(* IEC 61131-3 sources: daoli-st-library/DL_Base (part 20) *)

(* ---- FB_DL_PresetCounterSat.st ---- *)
(*==============================================================================
 * 组件名称 (Component)  : FB_DL_PresetCounterSat
 * 所属子库 (Sublibrary) : DL_Base
 * 当前版本 (Version)    : 1.0.1
 * 分类     (Category)   : 计数功能块（Function Block · Counter）
 * 兼容性   (Platform)   : CODESYS 3.5 / TwinCAT 3 / 汇川 InoProShop / Machine Expert
 *                         仅依赖 Standard.library（R_TRIG），零厂商方言
 * 功能简介 (Function)   : 带饱和预设计数器：上/下双向计数（上升沿生效），
 *                         到达上限（nPreset）或下限（nLowLimit）饱和不回绕
 *                         ——上计数在 nCount >= nPreset 时拒绝递增并保持
 *                         bSatHigh，下计数在 nCount <= nLowLimit 时拒绝递减
 *                         并保持 bSatLow。到达上限输出保持型完成标志 bDone
 *                         与单拍阈值事件 bThreshold（首次到达一拍脉冲，遵循
 *                         R25 单拍标志生命周期三律）。装载 bLoad 优先级最高，
 *                         复位 bReset 次之，同拍双计数互相抵消不偏置任何方向。
 *                         与已入库 FB_DL_EventCounter（回绕 + 比较输出通用
 *                         事件计数）、FB_DL_ModuloCounter（取模工位索引）
 *                         职责分离——本块是饱和计数（批次计数 / 托盘满载
 *                         场景），越界语义固定为钳位停走。
 * 开源溯源 (Origin)     : 原创实现（参考 LGF 库 Counter 计数器分类的功能域
 *                         与参数域，来源标签 lgf-counter），饱和计数语义为
 *                         公开计数器行为域，仅借分类/参数域/命名，clean-room
 *                         实现，未复制任何厂商私有库源码，不构成衍生作品。
 * 日期     (Date)       : 2026-11-15 ｜ 作者 (Author): Daoli Library
 * 依赖     (Depends)    : 无 DL_ 内部依赖；Standard.library: R_TRIG
 *
 *------------------------------------------------------------------------------
 * 【引脚契约 / Pin contract】
 *   输入 bCountUp   : BOOL — 上计数脉冲输入，上升沿 +1；
 *   输入 bCountDown : BOOL — 下计数脉冲输入，上升沿 -1；
 *   输入 bLoad      : BOOL — 装载预设值，上升沿生效（优先级最高）；
 *   输入 nPreset    : DINT — 上限预设值 [个]，>= nLowLimit，默认 100；
 *   输入 nLowLimit  : DINT — 下限预设值 [个]，<= nPreset，默认 0；
 *   输入 bReset     : BOOL — 复位到下限，上升沿生效（次优先级，兼故障解除）；
 *   输出 nCount     : DINT — 当前计数值 [个]，饱和域 [nLowLimit, nPreset]；
 *   输出 bSatHigh   : BOOL — 已达上限饱和（保持型，逐拍重算）；
 *   输出 bSatLow    : BOOL — 已达下限饱和（保持型，逐拍重算）；
 *   输出 bDone      : BOOL — 计数到达上限（保持型，逐拍重算）；
 *   输出 bThreshold : BOOL — 首次到达上限单拍脉冲（R25 三律）；
 *   输出 uErrorId   : UDINT — 故障码，0 = 无故障。
 *
 * 【优先级序 / Priority order（写死防歧义）】
 *   参数故障锁存 > 装载（bLoad 沿）> 复位（bReset 沿）> 同拍双计数抵消
 *   （计数值不变，不偏置任何方向）> 单向上计数 > 单向下计数 > 保持。
 *   同拍装载与计数脉冲：装载覆盖计数（计数脉冲被吞，不补发不记账）。
 *   同拍装载与复位：装载优先（覆盖复位到下限的行为）。
 *
 * 【饱和语义 / Saturation semantics（写死防误解）】
 *   上饱和：nCount = nPreset 时再收上计数沿 → 计数值保持 nPreset 不回绕、
 *           不取模，bSatHigh 保持 TRUE，脉冲被吞不置任何事件码（饱和本身
 *           是正常工况语义而非故障，上层以 bSatHigh/bDone 感知）；
 *   下饱和：nCount = nLowLimit 时再收下计数沿 → 保持 nLowLimit，bSatLow
 *           保持 TRUE，脉冲同样被吞；
 *   与 FB_DL_EventCounter 的 bWrap = FALSE 饱和模式语义一致但本块无回绕
 *   选项——批次/满载场景回绕是危险行为，设计上直接删除该自由度。
 *
 * 【bThreshold 单拍 R25 三律落地 / One-shot pulse lifecycle】
 *   置位律：仅「本拍到达上限 AND 上拍未在限」的扫描拍置 TRUE
 *           （bReached 为边沿基准，单一来源，仅由计数出口单点推导）；
 *   自清律：bThreshold 每拍预清 FALSE，无到达沿自动回落，不锁存；
 *   基准律：bReached 每拍在计数出口后单点刷新为 (nCount >= nPreset)，
 *           无第二份镜像状态；故障拍强制 bReached := FALSE，故障解除后
 *           再次到达会重新给出一拍脉冲（诊断链可见）。
 *
 * 【边界防错清单 / Boundary guard list】
 *   B1 nPreset < nLowLimit → 参数非法故障锁存 16#0001_0212：计数值强制钳到
 *      nLowLimit，计数/装载全部冻结，仅 bReset 上升沿解除（R15：故障级
 *      锁存仅解除路径清码）；解除后首次满足条件重新计数；
 *   B2 先判界后加减：上计数前判 nCount >= nPreset、下计数前判
 *      nCount <= nLowLimit，杜绝 DINT 极值 +1/-1 回绕穿透判据；
 *   B3 同拍 bCountUp/bCountDown 同时有效 → 计数不变（不偏置任何方向）；
 *   B4 装载值即 nPreset 引脚现值（装载拍实时采样，非缓存旧值）；
 *   B5 bReset 上升沿把计数值直接置 nLowLimit 并同时清除故障锁存。
 *
 * 【调用示例 / Call example】
 *   「托盘满载计数：装满 100 件给满托信号，人工换托后复位」
 *   fbPalletCnt(bCountUp := bPartInFeed, bCountDown := bPartRejectOut,
 *               bLoad := FALSE, nPreset := 100, nLowLimit := 0,
 *               bReset := bPalletChanged, nCount => nPalletCount,
 *               bSatHigh => , bSatLow => , bDone => bPalletFull,
 *               bThreshold => bPalletFullPulse, uErrorId => uCntErr);
 *
 * 【平台移植注意 / Porting notes】
 *   全部运算为 DINT 整数比较与加减，先判界后运算的次序保证永不触发
 *   DINT 极值回绕，无浮点、无除法、无定时依赖，各平台行为一致。
 *
 * 【工程背景与应用场景 / Background and use cases】
 *   ① 托盘满载计数：产线件流逐件 +1，装满 nPreset 件给满托信号（bDone/
 *      bThreshold），人工换托后 bReset 清零重新计件；
 *   ② 批次计数器：批次目标 nPreset 件，剔除品经 bCountDown 回退，计数
 *      上下饱和防止误键导致的负数或超量程静默错值；
 *   ③ 收线长度/圈数计量：到达设定圈数停机收卷（饱和停走保证计数器停在
 *      满值可读，回绕式计数会让操作工无法读出实际完成量）；
 *   ④ 重复触发防护：bThreshold 单拍脉冲驱动一次性动作（满托打印/批次
 *      结束报文），保持型 bDone 驱动持续状态（满托指示灯）。
 *
 * 【保持型与单拍输出关系表 / Held vs one-shot output relation】
 *   输出          类型     置位条件                     复位条件
 *   bSatHigh     保持型   nCount >= nPreset            nCount 降回限内
 *   bSatLow      保持型   nCount <= nLowLimit          nCount 升回限内
 *   bDone        保持型   nCount >= nPreset            nCount 降回限内/故障
 *   bThreshold   单拍     首次到达拍（含装载到达）      下一拍自动回落
 *   bSatHigh 与 bDone 判据相同但语义分层：bSatHigh 描述"在限停走状态"，
 *   bDone 描述"任务完成状态"，分开输出便于上层对停走与完成做不同联锁。
 *
 * 【典型时序推演 / Typical timing walkthrough】
 *   设 nPreset = 3，nLowLimit = 0，上电 nCount = 0：
 *     拍 1 上沿 → 1；拍 2 上沿 → 2；拍 3 上沿 → 3，bDone TRUE，
 *       bThreshold 单拍 TRUE，bSatHigh TRUE；
 *     拍 4 上沿 → 保持 3（上饱和），bThreshold FALSE（无新到达沿）；
 *     拍 5 下沿 → 2，bSatHigh/bDone 回落，bThreshold 无脉冲（2 不是到达）；
 *     拍 6 上沿 → 3，bThreshold 单拍 TRUE（bReached 已回落，重新到达）；
 *     拍 7 bReset 沿 → 0，bSatLow TRUE，无脉冲；
 *   结论：bThreshold 严格对应"从限外进入上限"的每一次跃迁，同限保持
 *   与复位不触发，装载到达触发（口径与验收推演 C1~C7 一致）。
 *
 * 【参数退化域 / Degenerate parameter domains】
 *   nPreset = nLowLimit：计数域退化为单点，装载到该点后双向均饱和停走
 *   （验收推演 C7）；上电 nCount = 0 若低于下限（如 nLowLimit = 5），
 *   bSatLow 立即为 TRUE，首个下计数沿被吞直至装载/复位对齐下限——
 *   上层应在上电后先装载或复位一次，保证计数值落在合法饱和域内。
 *
 * 【同族职责分离 / Family separation】
 *   FB_DL_EventCounter：通用事件计数（回绕/饱和双模式 + 阈值比较输出）；
 *   FB_DL_ModuloCounter：取模工位索引（循环工位场景）；本块：固定饱和
 *   计数（批次满载），三者语义正交、零互相调用。
 *
 * 红线自检 (Redline)    : R1 零全局变量表/外部变量引用 ✓ ｜ R2 零物理 IO 地址 ✓
 *                         R3 纯 IEC 61131-3 标准运算 ✓ ｜ R4 先判界后运算/
 *                           故障锁存仅解除路径清码/参数钳位 ✓
 *                         R5 全变量中英双语同行注释 ✓ ｜ R6 N/A（无主状态机，
 *                           优先级 IF-ELSIF 链即状态裁决，规格豁免 ENUM）✓
 *                         R7 四个 R_TRIG 主体最前部无条件刷新 ✓ ｜ R8 界限/
 *                           码值全常量化，无魔法数 ✓
 * 验收推演 (Acceptance) :
 *   C1 单发递增链：nPreset=3, nLowLimit=0，连发 3 个上沿 → 1/2/3，第 3 拍
 *      bDone TRUE 且 bThreshold 单拍 TRUE；第 4 个上沿 → 保持 3，bSatHigh
 *      TRUE，bThreshold 无脉冲；
 *   C2 下饱和：nCount=0 时发下沿 → 保持 0，bSatLow TRUE，无事件码；
 *   C3 同拍双计数：nCount=1 时同拍上/下沿 → 保持 1，无偏置；
 *   C4 装载优先：nCount=0 时同拍 bLoad 沿 + 上沿 → nCount := nPreset，
 *      bThreshold 单拍 TRUE（首次到达），上沿被覆盖不记账；
 *   C5 复位：bCount=5 时 bReset 沿 → nCount := nLowLimit，bDone/bSatHigh
 *      回落，bThreshold 无脉冲（复位不算"到达"）；
 *   C6 参数非法：nPreset=2 < nLowLimit=5 → 故障锁存 0212，nCount 强制 5，
 *      计数冻结；bReset 沿 → 当拍解除锁存并把计数压到下限，但同一拍段 3
 *      复检参数仍非法即刻**重新锁存**（参数不修正则计数不恢复）；须先把
 *      nPreset 改为 >= nLowLimit，再给 bReset 沿才彻底解除并可重新计数
 *      （v1.0.1 终审勘误：原文"bReset 沿 → 解除，可重新计数"未写明参数前置，
 *      与"锁存置位每拍检测"的实现不符）；
 *   C7 下限装载边界：nPreset = nLowLimit = 7 → 上电 nCount=0，bSatLow TRUE；
 *      bLoad 沿 → nCount := 7，bThreshold 单拍 TRUE，此后双向均饱和停走。
 *
 * 【故障码表 / Error code table】
 *   16#0001_0212  参数非法：上限预设 nPreset < 下限预设 nLowLimit，故障级
 *                 锁存，计数冻结在 nLowLimit，仅 bReset 上升沿解除（0212
 *                 空闲，0210/0211 已被 EventCounter/ModuloCounter 登记）。
 *
 * 【设计要点 / Key notes】
 *   ① 计数值单点出口：段 4 优先级链只写 nWork，段 4 末 nCount := nWork
 *      单点回写，故障段强制钳位也只改出口，任何路径不出现第二份计数镜像，
 *      杜绝多出口读改写竞态（沿用库内 EventCounter 修复后的单点出口范式）；
 *   ② 先判界后运算：加/减算全部在边界预判之后执行，DINT 极值 +1/-1 回绕
 *      在数学上不可达（R25 家族通用防穿透写法）；
 *   ③ 故障锁存生命周期：置位（段 3 每拍检测）→ 冻结（段 4 闸门）→ 解除
 *      （仅段 2 复位沿），三段各一入口，无第三条改动路径（R15）；
 *   ④ 饱和吞脉冲不置码：饱和属正常工况语义，置码会造成诊断链噪音，
 *      上层以 bSatHigh/bSatLow 感知（与 EventCounter 溢出一拍脉冲口径
 *      不同，两块语义分层，注释在两侧各自写死）；
 *   ⑤ 事件型组件免首扫：计数由脉冲沿驱动，无连续量同步语义，按 R23
 *      不设 bInit 跟踪逻辑，上电即处于下限饱和观测态。
 *
 * 【实现选择 / Implementation choice】
 *   无主状态机（规格豁免 ENUM）：饱和计数的行为本质是「边沿事件 + 优先级
 *   裁决 + 单点出口」，用 IF-ELSIF 优先级链表达比 ENUM+CASE 更短且无空态；
 *   计数值单点出口（nCount := _nWork 后全段共享），bSatHigh/bSatLow/bDone
 *   全部由出口值逐拍重算派生，无第二份计数镜像，杜绝读改写竞态；
 *   本块为事件型计数组件，无连续量同步语义，按 R23 免首扫，不设 bInit。
 *
 * 修订历史 (Revision)   :
 *   2026-11-15  v1.0.0  首版落盘（Round 09 · 泳道 A · LGF Counter 组）
 *   2026-11-15  v1.0.1  终审勘误：验收推演 C6 补写"参数未修正时 bReset 沿当拍
 *                       重新锁存"的前置条件（原文易误读为复位即可恢复计数）；
 *                       代码行为未改动，故障码 0001_0212 复核无冲突
 *============================================================================*)
FUNCTION_BLOCK FB_DL_PresetCounterSat
VAR_INPUT
    bCountUp   : BOOL;                     // 上计数脉冲输入，上升沿 +1 / Count-up pulse input, rising edge increments
    bCountDown : BOOL;                     // 下计数脉冲输入，上升沿 -1 / Count-down pulse input, rising edge decrements
    bLoad      : BOOL;                     // 装载预设值，上升沿生效（优先级最高）/ Load preset, rising edge, top priority
    nPreset    : DINT := 100;              // 上限预设值 [个]，>= nLowLimit / Upper preset [pieces], at least nLowLimit
    nLowLimit  : DINT := 0;                // 下限预设值 [个]，<= nPreset / Lower preset [pieces], at most nPreset
    bReset     : BOOL;                     // 复位到下限，上升沿生效（兼故障解除）/ Reset to lower limit, rising edge, also releases the fault latch
END_VAR
VAR_OUTPUT
    nCount     : DINT := 0;                // 当前计数值 [个]，饱和域 [nLowLimit, nPreset] / Current count [pieces], saturated within [nLowLimit, nPreset]
    bSatHigh   : BOOL;                     // 已达上限饱和（保持型）/ Saturated at upper limit (held)
    bSatLow    : BOOL;                     // 已达下限饱和（保持型）/ Saturated at lower limit (held)
    bDone      : BOOL;                     // 计数到达上限（保持型）/ Count reached upper limit (held)
    bThreshold : BOOL;                     // 首次到达上限单拍脉冲（R25 三律）/ First-arrival one-shot pulse (R25 three rules)
    uErrorId   : UDINT;                    // 故障码，0 = 无故障 / Error code, 0 = none
END_VAR
VAR
    fbTrigUp   : R_TRIG;                   // 上计数边沿 / Count-up edge detector
    fbTrigDn   : R_TRIG;                   // 下计数边沿 / Count-down edge detector
    fbTrigLoad : R_TRIG;                   // 装载边沿 / Load edge detector
    fbTrigRst  : R_TRIG;                   // 复位边沿 / Reset edge detector
    bReached   : BOOL := FALSE;            // 内部到达标志（阈值事件边沿基准，单一来源）/ Internal reached flag (threshold edge baseline, single source)
    bFaultLatch: BOOL;                     // 参数非法故障锁存（仅复位沿解除）/ Invalid-parameter fault latch (released only by reset edge)
    nWork      : DINT;                     // 计数运算工作副本（单点出口）/ Working copy for count arithmetic (single outlet)
    bUpEdge    : BOOL;                     // 本拍上计数沿有效 / Up edge active this scan
    bDnEdge    : BOOL;                     // 本拍下计数沿有效 / Down edge active this scan
    bLoadEdge  : BOOL;                     // 本拍装载沿有效 / Load edge active this scan
    bRstEdge   : BOOL;                     // 本拍复位沿有效 / Reset edge active this scan
END_VAR
VAR CONSTANT
    DL_CNT_ERR_PARAM : UDINT := 16#0001_0212; // 参数非法故障码（上限 < 下限）/ Error code for invalid parameters (preset below lower limit)
END_VAR

(*------------------------------------------------------------------------------
 * 段 1｜边沿实例无条件周期刷新（R7 红线：严禁置于 IF/CASE 分支内）
 *      Unconditional per-cycle refresh of all edge instances (R7 redline)
 *      四个 R_TRIG 全部在主体最前部刷新，与任何条件无关
 *      All four R_TRIG instances refreshed at the very top of the body
 *-----------------------------------------------------------------------------*)
fbTrigUp(CLK   := bCountUp);               // 上计数沿（Up edge）
fbTrigDn(CLK   := bCountDown);             // 下计数沿（Down edge）
fbTrigLoad(CLK := bLoad);                  // 装载沿（Load edge）
fbTrigRst(CLK  := bReset);                 // 复位沿（Reset edge）
bUpEdge   := fbTrigUp.Q;                   // 本拍上计数沿（Up edge this scan）
bDnEdge   := fbTrigDn.Q;                   // 本拍下计数沿（Down edge this scan）
bLoadEdge := fbTrigLoad.Q;                 // 本拍装载沿（Load edge this scan）
bRstEdge  := fbTrigRst.Q;                  // 本拍复位沿（Reset edge this scan）

(*------------------------------------------------------------------------------
 * 段 2｜输出预清零（R25 自清律）+ 复位/故障解除路径
 *      Output preset clearing (R25 self-clear rule) + reset/release paths
 *      bThreshold 每拍预清 FALSE：无到达沿自动回落，不锁存
 *      bThreshold preset FALSE each scan: falls back without an arrival edge
 *-----------------------------------------------------------------------------*)
bThreshold := FALSE;                       // 单拍脉冲预清（One-shot preset cleared）
uErrorId   := 16#0000_0000;                // 故障码出口预清，段 6 按锁存态重写 / Error outlet preset, rewritten by stage 6 per latch state

IF bRstEdge THEN                           // 复位沿：计数回下限并解除故障锁存 / Reset edge: count back to lower limit and release the latch
    bFaultLatch := FALSE;                  // 故障锁存解除（R15 解除路径唯一）/ Latch released (unique release path per R15)
    nWork       := nLowLimit;              // 计数值回下限（Count back to lower limit）
    nCount      := nWork;                  // 计数单点出口（Single outlet）
END_IF

(*------------------------------------------------------------------------------
 * 段 3｜参数防御（边界 B1）：nPreset < nLowLimit → 故障锁存，计数冻结
 *      Parameter guard (B1): preset below lower limit latches a fault
 *   锁存期间计数值强制钳到 nLowLimit、全部计数/装载动作冻结，仅复位沿解除
 *   While latched, count is forced to nLowLimit and all actions frozen
 *   锁存生命周期三段：置位（本段检测）→ 冻结（段 4 闸门跳过）→ 解除（段 2
 *   复位沿），每段单入口，无第三条改动路径（R15 故障级公约）
 *   Latch lifecycle: raise here, freeze in stage 4, release only in stage 2
 *-----------------------------------------------------------------------------*)
IF nPreset < nLowLimit THEN
    bFaultLatch := TRUE;                    // 参数非法故障锁存（Invalid-parameter latch）
END_IF

IF NOT bFaultLatch THEN

    (*--------------------------------------------------------------------------
     * 段 4｜计数主逻辑（优先级序写死）：装载 > 复位 > 双计数抵消 > 单向
     *      Counting main logic (fixed priority): load > reset > cancel > single
     *   注意复位沿已在段 2 处理计数值回下限，此处 ELSIF 链只在非复位拍进入；
     *   同拍装载与复位冲突时装载胜出（覆盖段 2 的回下限值）
     *   A load edge on the same scan as reset wins over the reset value
     *-------------------------------------------------------------------------*)
    IF bLoadEdge THEN
        nWork := nPreset;                   // 装载优先级最高：写入引脚现值（Load top priority: live pin value）
    ELSIF bRstEdge THEN
        nWork := nLowLimit;                 // 复位次之：回到下限（Reset next: back to lower limit）
    ELSIF bUpEdge AND bDnEdge THEN
        nWork := nCount;                    // 同拍双计数抵消：计数不变不偏置（Dual edges cancel: no bias）
        (* 口径注释：双沿抵消不置事件码——抵消属输入侧拍点重叠的正常现象，
           置码会造成诊断噪音；与 EventCounter 的信息级 0101 抵消码口径
           不同（该块有显式抵消码），本块按规格只保证"不偏置任何方向" *)
    ELSIF bUpEdge THEN
        IF nCount >= nPreset THEN
            nWork := nPreset;               // 上饱和：钳位停走不回绕（Upper saturation: clamp and hold, no wrap）
        ELSE
            nWork := nCount + 1;            // 先判界后加算，无极值回绕（Boundary pre-checked increment）
        END_IF
    ELSIF bDnEdge THEN
        IF nCount <= nLowLimit THEN
            nWork := nLowLimit;             // 下饱和：钳位停走不回绕（Lower saturation: clamp and hold, no wrap）
        ELSE
            nWork := nCount - 1;            // 先判界后减算，无极值回绕（Boundary pre-checked decrement）
        END_IF
    ELSE
        nWork := nCount;                    // 无事件保持（No event, hold）
    END_IF
    nCount := nWork;                        // 计数单点出口（Single outlet for the count）
END_IF

(*------------------------------------------------------------------------------
 * 段 5｜保持型输出派生：全部由计数出口逐拍重算，无第二份镜像
 *      Held outputs derived from the count outlet each scan, no mirror state
 *   派生式而非锁存式：三路保持型输出每拍从计数出口现值重算，即使计数
 *   被装载/复位/故障强行搬移，输出也在同拍对齐，无跨拍错位窗口；
 *   bSatHigh 与 bDone 判据相同但语义分层（停走态 vs 完成态），见头注释
 *   关系表，上层可分别做联锁与指示。
 *-----------------------------------------------------------------------------*)
IF bFaultLatch THEN
    nCount   := nLowLimit;                  // 故障期计数值强制钳到下限（Forced clamp while latched）
    bSatHigh := FALSE;                      // 故障期上限饱和态清空（Upper saturation cleared while latched）
    bSatLow  := TRUE;                       // 故障期钳在下限 → 下饱和态成立（Clamped at lower limit, so lower saturation holds）
    bDone    := FALSE;                      // 故障期完成标志清空（Done cleared while latched）
ELSE
    bSatHigh := (nCount >= nPreset);        // 上饱和派生（Upper saturation derived）
    bSatLow  := (nCount <= nLowLimit);      // 下饱和派生（Lower saturation derived）
    bDone    := (nCount >= nPreset);        // 完成标志派生（Done derived）
END_IF

(*------------------------------------------------------------------------------
 * 段 6｜bThreshold 单拍脉冲（R25 三律：置位/自清/基准单一来源）
 *      bThreshold one-shot pulse (R25: set / self-clear / single-source baseline)
 *   置位：本拍在限 AND 上拍未在限（bReached 边沿基准）；
 *   自清：段 2 每拍预清，无沿自动回落；
 *   基准：bReached 本拍末单点刷新，故障拍强制 FALSE（解除后可再触发）。
 *   装载/计数任一路径到达上限均视为"到达"（口径写死）；
 *   复位路径回下限不算到达，不给脉冲（验收推演 C5）。
 *   跃迁真值表（上拍 bReached → 本拍在限 → bThreshold）：
 *     FALSE → TRUE  ：单拍 TRUE（首次到达或离开后重新到达）
 *     TRUE  → TRUE  ：FALSE（同限保持不触发）
 *     任意  → FALSE ：FALSE（离开上限不触发，下限侧无阈值事件）
 *-----------------------------------------------------------------------------*)
IF (NOT bFaultLatch) AND (nCount >= nPreset) AND (NOT bReached) THEN
    bThreshold := TRUE;                     // 首次到达单拍脉冲（First-arrival one-shot）
END_IF

IF bFaultLatch THEN
    bReached := FALSE;                      // 故障拍强制清基准，解除后可再触发 / Baseline force-cleared while latched, re-armable after release
ELSE
    bReached := (nCount >= nPreset);        // 边沿基准单点刷新（Baseline refreshed at a single point）
END_IF

(*------------------------------------------------------------------------------
 * 段 7｜uErrorId 出口（R15：故障级锁存优先透出）
 *      uErrorId outlet (R15: latched fault code has priority)
 *-----------------------------------------------------------------------------*)
IF bFaultLatch THEN
    uErrorId := DL_CNT_ERR_PARAM;           // 参数非法锁存码（Latched parameter code）
ELSE
    uErrorId := 16#0000_0000;               // 无故障透出零码（Zero when healthy）
END_IF

(*------------------------------------------------------------------------------
 * 段 8｜验收推演索引 / Acceptance walkthrough index
 *   C1 递增链 1/2/3 → 第 3 拍 bDone+单拍；第 4 拍饱和停走无脉冲
 *   C2 下饱和保持 0；C3 双沿抵消不偏置；C4 装载覆盖计数并给单拍
 *   C5 复位回下限无脉冲；C6 参数非法锁存 0212 仅复位沿解除
 *   C7 nPreset = nLowLimit 退化域：装载拍单拍触发后双向饱和
 *-----------------------------------------------------------------------------*)
END_FUNCTION_BLOCK

(* ---- FB_DL_RolloverCounter.st ---- *)
(*==============================================================================
 * 组件名称 (Component)  : FB_DL_RolloverCounter
 * 所属子库 (Sublibrary) : DL_Base
 * 当前版本 (Version)    : 1.0.0
 * 分类     (Category)   : 计数功能块（Function Block · Counter）
 * 兼容性   (Platform)   : CODESYS 3.5 / TwinCAT 3 / 汇川 InoProShop / Machine Expert
 *                         仅依赖 Standard.library（R_TRIG / MIN），零厂商方言
 * 功能简介 (Function)   : 回绕型可逆计数器。在 0 至回绕上限的环形域内上下计数，
 *                         到顶继续加则回 0、到底继续减则回上限，同时输出回绕单拍
 *                         脉冲与**净回绕圈数**（可负），用于转盘圈数统计、编码器
 *                         溢出圈数、料盘循环计数等「只关心绕了多少圈」的场合。
 *                         本块**不做任何预设比较逻辑**：既不在到达预设时冻结，
 *                         也不做双预设区间判断，纯粹计数 + 回绕 + 圈数累积。
 *
 * 【引脚契约 / Pin contract】
 *   输入 bEnable      : BOOL  — 使能。FALSE 时冻结计数（值保持、圈数保持、无脉冲），
 *                               状态回空闲；本块不因失能清零，清零只认复位沿；
 *   输入 bReset       : BOOL  — 上升沿把计数值与圈数清零（可在任意状态生效）；
 *   输入 bCountUp     : BOOL  — 上升沿加计数（电平保持不重复计数）；
 *   输入 bCountDown   : BOOL  — 上升沿减计数（电平保持不重复计数）；
 *   输入 bLoad        : BOOL  — 电平有效装载，优先级最高（高于复位沿与计数沿）；
 *   输入 uLoadValue   : UDINT — 装载值 [cnt]，超过回绕上限时钳位并置信息码；
 *   输入 uPreset      : UDINT — 回绕上限（含）[cnt]，有效域 1~16#FFFF_FFFE；
 *   输出 uCount       : UDINT — 当前计数值 [cnt]，0 ~ 回绕上限；
 *   输出 bWrapped     : BOOL  — 本拍发生回绕的单拍脉冲（上下回绕均置位）；
 *   输出 nTurns       : DINT  — 净回绕圈数 [圈]，上加下减，可负，带饱和保护；
 *   输出 bAtPreset    : BOOL  — 当前值已达回绕上限（逐拍重算，非锁存）；
 *   输出 eState       : ENUM  — 主状态机当前态（E_DL_RolloverPhase）；
 *   输出 bError       : BOOL  — 故障锁存：回绕上限退化（小于 1），计数冻结；
 *   输出 uErrorId     : UDINT — 事件 / 故障码，0 = 无。
 *
 * 【与既有四件计数器的职责边界 / Family separation（五件互斥，写死不可互替）】
 *   FB_DL_EventCounter         = 单向事件累加（只关心总数）；
 *   FB_DL_ModuloCounter        = 取模工位索引（单向，用取模得余数）；
 *   FB_DL_PresetCounterSat     = 单向双预设饱和（到限冻结，不回绕）；
 *   FB_DL_BidirectionalCounter = CTUD 双预设比较（关心区间高低限）；
 *   本块                       = 环形回绕 + 净圈数（无预设比较，只关心绕圈）。
 *   本块刻意不实现「到限冻结」与「取模」：前者是饱和件语义，后者在无符号域与
 *   有符号域上行为不一致（历史坑），本块回绕一律用「比较 + 赋值」实现，禁 MOD。
 *
 * 【计数优先级 / Priority chain（同拍多指令的仲裁口径）】
 *   ① 回绕上限退化（小于 1）→ 冻结，最高优先级，任何计数沿都不生效；
 *   ② 装载（bLoad 电平有效）→ 覆盖计数，同拍计数沿被丢弃；
 *   ③ 复位沿 → 计数与圈数清零（与装载同拍时装载胜出，因装载在其后执行）；
 *   ④ 双向同拍 → 净变化 0，计数不变、不发脉冲、置信息码 0120；
 *   ⑤ 单向沿 → 加 / 减，跨过上下界即回绕并累计圈数。
 *
 * 【指令优先级矩阵 / Priority matrix（行 = 状态，列 = 本拍指令）】
 *   状态 \ 指令        退化   装载   复位沿   双向同拍   单向上/下   无指令
 *   eIdle              冻结   落计数 清零     落计数     落计数      保持
 *   eCount             冻结   装载     清零     丢弃       加减回绕    保持
 *   eFrozen            保持   保持     退出冻结 保持       保持        保持
 *   矩阵口径写死：装载是「电平」而非沿，保持期间每拍都写同一个值；
 *   复位是「沿」，只在上升沿那一拍动作；计数同样只认沿，电平保持不重复计数。
 *   三者混用时按上表逐格落地，不存在「装载与计数同拍谁先谁后」的解释空间。
 *
 * 【回绕与圈数口径 / Wrap and turn semantics】
 *   加法回绕：当前值已达上限（大于等于上限）→ 计数值回 0，圈数 +1；
 *   减法回绕：当前值为 0 → 计数值回上限，圈数 -1；
 *   圈数饱和：nTurns 触及正 / 负饱和上限后停在该值，并置信息码（不再累加），
 *   防止远端诊断页数值溢出翻转（历史 D 类缺陷）。饱和后需复位沿才能重新累计。
 *
 * 【圈数换算与量程校核 / Turn-to-engineering conversion】
 *   真实位移 = nTurns × 一圈当量 + 当前值 × 单格当量（一圈当量 = 上限 + 1 格）；
 *   例：分度盘 60 格、单格 6 度，则 nTurns × 360 + uCount × 6 即累计角度；
 *   量程校核方法：nTurns 饱和值 2×10^9 圈 × 一圈当量，须仍在调用方量程内，
 *   量程不足时调用方应在换向或换批时用复位沿清零，而不是依赖饱和兜底。
 *   本块输出「净圈数」而非「绝对位置」：掉电重启后圈数从 0 起算，
 *   需要绝对位置时由调用方在上电时用装载引脚把已知位置写入并自行保存圈数。
 *
 * 【饱和与复位的配合 / Saturation versus reset】
 *   饱和只是停止累加，不改写任何已有值：回绕脉冲照发、计数值照转，
 *   因此「绕圈事实」不会因为圈数饱和而丢失，只是不再累进到诊断量上；
 *   复位沿同时清零计数与圈数并解除饱和，是唯一的重入手段；
 *   本块不因使能撤除而清零：失能只冻结，避免产线短暂停机就丢失圈数。
 *
 * 【现场整定与故障定位提示 / Commissioning hints】
 *   ① 上电先给一次复位沿，把计数与圈数拉到已知零点，再开始累计；
 *   ② 空载手转一圈，观察 bWrapped 是否恰好出现一次：出现两次说明上限设小了，
 *      一次都不出现说明上限大于实际一圈格数（脉冲被吃掉）；
 *   ③ 计数跳变排查：若 uCount 出现跨格跳跃，先查引脚注入的脉冲是否被上层
 *      做了防抖（防抖会削沿，本块只认沿，不做任何滤波）；
 *   ④ 圈数与机械圈数不符时，优先核对上限是否为「一圈格数减一」（上限含端点）。
 *
 * 【主状态机 / Main state machine（ENUM + CASE + ELSE 兜底）】
 *   eIdle   → bEnable 且上限合法：eCount；
 *   eIdle   → bEnable 但上限退化：eFrozen 并置 0218；
 *   eCount  → 上限退化：eFrozen（计数保持，不回 0，避免死循环式跳动）；
 *   eCount  → 使能撤除：eIdle（计数冻结保持）；复位沿留在 eCount 内清零；
 *   eFrozen → 上限恢复合法或复位沿：eIdle（复位后重新装载）；
 *   eFrozen → 使能撤除：eIdle；
 *   ELSE    → 非法态值：eFrozen 并置 0218（兜底拦截，绝不落空态）。
 *
 * 【边界防错清单 / Boundary guard list】
 *   B1 回绕上限小于 1（含 0）→ 退化冻结：不回绕到 0、不产生无穷回绕，置 0218；
 *   B2 回绕上限超过 16#FFFF_FFFE → 钳到该值并置 0120（防极端值参与比较歧义）；
 *   B3 装载值超上限 → 钳到上限并置 0120（钳位后仍接受装载，不丢弃指令）；
 *   B4 双向同拍 → 计数不变、脉冲不发、置 0120（避免扫描时序歧义）；
 *   B5 圈数饱和 → 停在 ±饱和值并置 0120，不静默回绕；
 *   B6 整数域全为无符号 / 有符号整数比较（UDINT / DINT），无浮点参与，
 *      浮点判等容差红线在本块不适用（头注释显式声明）；
 *   B7 加法不做「上限 + 1」运算、减法不做「0 - 1」运算：回绕由直接赋值完成，
 *      无符号下溢 / 上溢永不发生，跨平台无差异。
 *
 * 【单拍标志三律 / One-shot pulse lifecycle（R24 / R25）】
 *   置位律：bWrapped 每拍于段 1 预清 FALSE，仅由段 5 的回绕分支置位；
 *   分离律：边沿「消费」在段 2 的实例 Q，脉冲「转出」在段 5 的计数分支，
 *           下一拍由段 1 预清零自清，不存在跨拍悬挂；
 *   基准律：三个边沿实例固定在主体顶层无条件刷新，基准唯一（引脚电平），
 *           不置于条件分支内，扫描抖动不丢沿、不重沿。
 *
 * 【调用示例 / Call example（仅行注释，不嵌套块注释）】
 *   // 分度盘：每工位 1 个脉冲，60 工位一圈，统计已转圈数与每圈回绕沿
 *   // fbTurn(fbIndex(bEnable := bRunOk, bReset := bIdxReset,
 *   //        bCountUp := bStationPulse, bCountDown := FALSE,
 *   //        bLoad := bHomingDone, uLoadValue := uHomePos, uPreset := 59,
 *   //        uCount => uStationNo, bWrapped => bLapDone,
 *   //        nTurns => nLapCount, bAtPreset => bLastStation,
 *   //        eState => eTurnState, bError => bTurnErr, uErrorId => uTurnErrId));
 *
 * 【平台移植注意 / Porting notes】
 *   UDINT 的比较与赋值在三平台语义一致；本块不使用 MOD 与无符号减法下溢，
 *   因此不存在「无符号回绕到 4294967295」这一类平台差异；DINT 饱和判据用
 *   显式比较而非加减后判溢出，避免依赖溢出标志位（部分平台不暴露该标志）。
 *
 * 【工程背景与应用场景 / Background and use cases】
 *   ① 分度盘 / 转盘：工位脉冲计数到一圈末回绕，回绕沿驱动「整圈完成」逻辑；
 *   ② 编码器 / 计量轮：增量计数的绝对值溢出后回绕，圈数用于累计真实行程；
 *   ③ 料盘循环：料盘码位循环取料，回绕沿触发一次空盘检测；
 *   ④ 卷绕 / 收放卷：正反转计数，净圈数直接反映卷径变化趋势（配合卷径计算件）。
 *
 * 【与上层逻辑的组合契约 / Composition contract】
 *   本块只做「环形计数 + 圈数」，不含任何工艺判断，也不输出报警级别；
 *   上层典型组合：
 *     回绕脉冲 → 触发「整圈完成」事务（发一次 HMI 计米更新或一次换盘请求）；
 *     到限标志 → 作为「下一格即回绕」的预判，供减速 / 预动作使用；
 *     圈数 + 计数 → 由上层换算为长度、角度或位置，本块不做量纲换算；
 *     故障位 → 并入设备级诊断汇总，本块不直接驱动任何硬件输出。
 *   本块不持有任何外部实体引用，也不回调上层：只有引脚进、引脚出。
 *
 * 【典型时序推演 / Typical timing walkthrough】
 *   设上限 100、初始计数 98：加沿 → 99；加沿 → 100（bAtPreset TRUE、无脉冲）；
 *   再加沿 → 计数 0、bWrapped 单拍 TRUE、圈数 +1；此后再加沿回常规递增。
 *   减向：计数 0 时减沿 → 计数 100、bWrapped 单拍 TRUE、圈数 -1。
 *   装载：bLoad 保持 TRUE 期间每拍把装载值写入计数，脉冲不产生；
 *   装载撤销后从装载值继续，圈数不变（装载不重置圈数，只有复位沿才清圈数）。
 *
 * 【验收向量 / Acceptance vectors】
 *   V1 上回绕：上限 100、计数 100、加沿 → 计数 0、bWrapped TRUE、圈数 +1；
 *   V2 下回绕：计数 0、减沿 → 计数 100、bWrapped TRUE、圈数 -1；
 *   V3 装载优先：bLoad TRUE、装载值 42、同拍有加沿 → 计数 42、圈数不变、无脉冲；
 *   V4 双向冲突：加沿与减沿同拍 → 计数不变、无脉冲、uErrorId 0120；
 *   V5 上限退化：上限 0、连续给加沿 → 计数保持、bError TRUE、uErrorId 0218。
 *   V6 装载钳位：上限 100、装载值 500、bLoad TRUE → 计数 100、uErrorId 0120；
 *   V7 连续绕圈：上限 9、从 0 起连给 30 个加沿 → 计数 0、圈数 +3、脉冲仅三次；
 *   V8 复位清圈：任意圈数下给一次复位沿 → 计数 0、圈数 0、脉冲不发。
 *
 * 【故障码表 / Error code table】
 *   16#0001_0120  信息级：装载值超上限已钳位 / 上下限超域已钳位 /
 *                 同拍双向已丢弃 / 圈数饱和已停止累加，均只进事件码；
 *   16#0001_0218  故障级：回绕上限小于 1（退化），计数冻结并锁存 bError。
 *
 * 修订历史 (Revision)   :
 *   2026-11-15  v1.0.0  首版落盘（Round 11 · 泳道 A · LGF Counter 组）
 *
 * 同文件发布类型 (Co-published type) : E_DL_RolloverPhase（本块主状态机枚举，
 *   按库内惯例随宿主 POU 同文件发布，禁止在其他文件重复声明同名枚举）。
 *============================================================================*)
TYPE E_DL_RolloverPhase :
(
    eIdle   := 0,      // 空闲：未使能，计数与圈数保持 / Idle, disabled, count and turns held
    eCount  := 10,     // 计数：按边沿加减并回绕 / Counting, edge driven with wrap-around
    eFrozen := 20      // 冻结：上限退化，计数保持且报警 / Frozen, degenerate bound, count held
);
END_TYPE

FUNCTION_BLOCK FB_DL_RolloverCounter
VAR_INPUT
    bEnable      : BOOL;                   // 使能，FALSE 时冻结计数 / Enable, FALSE freezes the counting
    bReset       : BOOL;                   // 上升沿清零计数与圈数 / Rising edge clears the count and the turns
    bCountUp     : BOOL;                   // 上升沿加计数 / Rising edge increments
    bCountDown   : BOOL;                   // 上升沿减计数 / Rising edge decrements
    bLoad        : BOOL;                   // 电平有效装载，优先级最高 / Level-true load, highest priority
    uLoadValue   : UDINT;                  // 装载值 [cnt]，超上限时钳位 / Load value [cnt], clamped to the bound
    uPreset      : UDINT;                  // 回绕上限（含）[cnt]，1~16#FFFF_FFFE / Wrap bound inclusive [cnt], 1 to 16#FFFF_FFFE
END_VAR
VAR_OUTPUT
    uCount       : UDINT;                  // 当前计数值 [cnt]，0 ~ 上限 / Current count [cnt], 0 to the bound
    bWrapped     : BOOL;                   // 本拍回绕单拍脉冲 / One-shot wrap pulse of this scan
    nTurns       : DINT;                   // 净回绕圈数 [圈]，上加下减 / Net wrap turns [turn], signed
    bAtPreset    : BOOL;                   // 当前值已达上限 / The count reached the bound
    eState       : E_DL_RolloverPhase;     // 主状态机当前态 / Current state of the main state machine
    bError       : BOOL;                   // 故障锁存：上限退化 / Fault latched, degenerate bound
    uErrorId     : UDINT;                  // 事件 / 故障码，0 = 无 / Event or fault code, 0 = none
END_VAR
VAR
    _eState      : E_DL_RolloverPhase;     // 内部状态寄存器，段 6 为唯一写点 / Internal state register, single writer in stage 6
    _fbTrigUp    : R_TRIG;                 // 加计数上升沿实例，顶层无条件刷新 / Rising-edge instance of the up pulse
    _fbTrigDown  : R_TRIG;                 // 减计数上升沿实例，顶层无条件刷新 / Rising-edge instance of the down pulse
    _fbTrigReset : R_TRIG;                 // 复位上升沿实例，顶层无条件刷新 / Rising-edge instance of the reset pin
    _uBound      : UDINT;                  // 钳位后的回绕上限工作副本 [cnt] / Working copy of the clamped bound [cnt]
    _bBoundOk    : BOOL;                   // 上限合法性标志 / Bound validity flag
    _bUpEdge     : BOOL;                   // 本拍加沿有效 / Up edge active in this scan
    _bDownEdge   : BOOL;                   // 本拍减沿有效 / Down edge active in this scan
    _bResetEdge  : BOOL;                   // 本拍复位沿有效 / Reset edge active in this scan
    _bWrapNow    : BOOL;                   // 本拍回绕已发生（消费拍标志）/ Wrap happened in this scan, consumer flag
    _nTurnStep   : DINT;                   // 本拍圈数增量 [圈]，+1 / -1 / 0 / Turn increment of this scan [turn]
END_VAR
VAR CONSTANT
    DL_PRESET_MIN : UDINT := 1;            // 上限下限 [cnt]，小于它即退化 / Lower bound of the wrap bound [cnt]
    DL_PRESET_MAX : UDINT := 16#FFFF_FFFE; // 上限上界 [cnt]，极端值参与比较易生歧义 / Upper bound of the wrap bound [cnt]
    DL_TURNS_MAX  : DINT  := 2000000000;   // 圈数饱和上限 [圈]，留累加余量 / Turn saturation limit [turn], leaves headroom
    DL_TURN_UP    : DINT  := 1;            // 圈数增量：加向回绕 [圈] / Turn increment for an up wrap [turn]
    DL_TURN_DOWN  : DINT  := -1;           // 圈数增量：减向回绕 [圈] / Turn increment for a down wrap [turn]
    DL_TURN_HOLD  : DINT  := 0;            // 圈数增量：不回绕 [圈] / Turn increment when no wrap occurs [turn]
    DL_ERR_INFO   : UDINT := 16#0001_0120; // 信息级码：钳位 / 冲突 / 饱和 / Info code for clamp, conflict and saturation
    DL_ERR_PRESET : UDINT := 16#0001_0218; // 故障级码：上限退化，计数冻结 / Fault code for a degenerate bound
END_VAR

(*------------------------------------------------------------------------------
 * 段 1｜输出与工作标志预清零（单拍标志置位律的起点）
 *      Preset clearing of outputs and working flags
 *   uCount / nTurns / bError 为跨拍保持量，此处不清；bWrapped 必须每拍预清。
 *-----------------------------------------------------------------------------*)
bWrapped   := FALSE;                       // 回绕脉冲预清（Wrap pulse preset）
bAtPreset  := FALSE;                       // 到限标志预清（Bound-reached flag preset）
uErrorId   := 16#0000_0000;                // 事件码预清零，逐段置位（Event code preset to zero）
_bWrapNow  := FALSE;                       // 回绕消费标志预清（Wrap consumer flag preset）
_nTurnStep := DL_TURN_HOLD;                // 圈数增量预置 0（Turn increment preset to zero）

(*------------------------------------------------------------------------------
 * 段 2｜边沿实例无条件周期刷新（周期安全红线）
 *      Unconditional per-cycle refresh of all edge instances
 *   三个实例固定在主体顶层，严禁挪入 IF / CASE 分支，否则边沿丢失、计数丢拍。
 *-----------------------------------------------------------------------------*)
_fbTrigUp(CLK    := bCountUp);             // 加计数上升沿（Increment rising edge）
_fbTrigDown(CLK  := bCountDown);           // 减计数上升沿（Decrement rising edge）
_fbTrigReset(CLK := bReset);               // 复位上升沿（Reset rising edge）

_bUpEdge    := _fbTrigUp.Q;               // 本拍加沿（Up edge of this scan）
_bDownEdge  := _fbTrigDown.Q;             // 本拍减沿（Down edge of this scan）
_bResetEdge := _fbTrigReset.Q;            // 本拍复位沿（Reset edge of this scan）

(*------------------------------------------------------------------------------
 * 段 3｜上限钳位与合法性判定（边界 B1 / B2）
 *      Bound clamping and validity verdict
 *   上界超域先钳位（防极端值参与比较），下界退化只判不钳：
 *   退化必须冻结而不是悄悄改成 1，否则现场永远看不到组态错误。
 *-----------------------------------------------------------------------------*)
_uBound := uPreset;                        // 上限工作副本接管输入（Bound working copy）
IF _uBound > DL_PRESET_MAX THEN            // 超上界（Above the upper bound）
    _uBound  := DL_PRESET_MAX;             // 钳到上界（Clamp to the upper bound）
    uErrorId := DL_ERR_INFO;               // 置钳位信息码（Raise the clamp info code）
END_IF

IF _uBound < DL_PRESET_MIN THEN            // 低于下限，退化（Below the lower bound, degenerate）
    _bBoundOk := FALSE;                    // 上限不可用（Bound unusable）
    bError    := TRUE;                     // 故障锁存（Latch the fault）
    uErrorId  := DL_ERR_PRESET;            // 置退化故障码（Raise the degenerate fault code）
ELSE                                       // 上限可用（Bound usable）
    _bBoundOk := TRUE;                     // 上限合法（Bound valid）
    bError    := FALSE;                    // 条件解除即清故障（Fault clears once the condition is gone）
END_IF

(*------------------------------------------------------------------------------
 * 段 4｜复位段（计数与圈数清零，任意状态生效）
 *      Reset stage, effective in every state
 *   复位在装载之前执行：同拍既复位又装载时装载胜出（装载语义为「强制落到某值」）。
 *-----------------------------------------------------------------------------*)
IF _bResetEdge THEN                        // 复位沿（Reset edge）
    uCount  := 0;                          // 计数清零（Count cleared）
    nTurns  := 0;                          // 圈数清零（Turns cleared）
    bWrapped := FALSE;                     // 同拍不发回绕脉冲（No wrap pulse on the reset scan）
END_IF

(*------------------------------------------------------------------------------
 * 段 5｜主状态机与计数核心（ENUM + CASE + ELSE 兜底）
 *      Main state machine with the counting core
 *   状态迁移与计数动作在同一 CASE 内完成，状态寄存器只有本段一个写点；
 *   回绕动作只在 eCount 分支里出现，退化态与空闲态不产生任何回绕。
 *-----------------------------------------------------------------------------*)
CASE _eState OF

    E_DL_RolloverPhase.eIdle:              // 空闲：等待使能（Idle, waiting for enable）
        IF bEnable AND _bBoundOk THEN      // 使能且上限合法（Enabled with a valid bound）
            _eState := E_DL_RolloverPhase.eCount;            // 进入计数态（Enter the counting state）
        ELSIF bEnable THEN                 // 使能但上限退化（Enabled but the bound is degenerate）
            _eState := E_DL_RolloverPhase.eFrozen;           // 进入冻结态（Enter the frozen state）
            uErrorId := DL_ERR_PRESET;     // 置退化故障码（Raise the degenerate fault code）
        END_IF

    E_DL_RolloverPhase.eCount:             // 计数：按优先级链处理本拍指令（Counting with the priority chain）
        IF NOT _bBoundOk THEN              // 上限转退化（The bound became degenerate）
            _eState  := E_DL_RolloverPhase.eFrozen;          // 进入冻结态，计数保持（Frozen, count held）
            uErrorId := DL_ERR_PRESET;     // 置退化故障码（Raise the degenerate fault code）
        ELSIF NOT bEnable THEN             // 使能撤除（Enable removed）
            _eState := E_DL_RolloverPhase.eIdle;             // 回空闲，计数冻结（Back to idle, count frozen）
        ELSIF bLoad THEN                   // 装载优先，电平有效（Load has the highest priority）
            IF uLoadValue > _uBound THEN   // 装载值超上限（Load value above the bound）
                uCount   := _uBound;       // 钳到上限（Clamp to the bound）
                uErrorId := DL_ERR_INFO;   // 置钳位信息码（Raise the clamp info code）
            ELSE                           // 装载值在域内（Load value within range）
                uCount := uLoadValue;      // 直接装载（Take the load value as-is）
            END_IF
            bWrapped := FALSE;             // 装载拍不发回绕脉冲（No wrap pulse on a load scan）
        ELSIF _bUpEdge AND _bDownEdge THEN // 双向同拍（Both edges in the same scan）
            uErrorId := DL_ERR_INFO;       // 方向冲突已丢弃（Direction conflict discarded）
        ELSIF _bUpEdge AND (NOT _bResetEdge) THEN  // 加向，复位拍不重复加减（Increment, skipped on a reset scan）
            IF uCount >= _uBound THEN      // 已达上限，触发上回绕（At the bound, wrap upwards）
                uCount    := 0;            // 回绕到 0（Wrap to zero）
                _bWrapNow := TRUE;         // 标记本拍回绕（Flag the wrap of this scan）
                _nTurnStep := DL_TURN_UP;  // 圈数增量 +1（Turn increment plus one）
            ELSE                           // 未到上限（Below the bound）
                uCount := uCount + 1;      // 常规加 1（Plain increment）
                _nTurnStep := DL_TURN_HOLD;// 圈数不变（Turns unchanged）
            END_IF
        ELSIF _bDownEdge AND (NOT _bResetEdge) THEN  // 减向，复位拍不重复加减（Decrement, skipped on a reset scan）
            IF uCount = 0 THEN             // 已在下界，触发下回绕（At zero, wrap downwards）
                uCount    := _uBound;      // 回绕到上限（Wrap to the bound）
                _bWrapNow := TRUE;         // 标记本拍回绕（Flag the wrap of this scan）
                _nTurnStep := DL_TURN_DOWN;// 圈数增量 -1（Turn increment minus one）
            ELSE                           // 未到下界（Above zero）
                uCount := uCount - 1;      // 常规减 1（Plain decrement）
                _nTurnStep := DL_TURN_HOLD;// 圈数不变（Turns unchanged）
            END_IF
        END_IF

    E_DL_RolloverPhase.eFrozen:            // 冻结：上限退化，计数保持（Frozen, count held）
        IF NOT bEnable THEN                // 使能撤除（Enable removed）
            _eState := E_DL_RolloverPhase.eIdle;             // 回空闲（Back to idle）
        ELSIF _bBoundOk THEN               // 组态已修正（Configuration fixed）
            _eState := E_DL_RolloverPhase.eIdle;             // 回空闲后重新装载（Back to idle, then re-enter counting）
        ELSIF _bResetEdge THEN             // 复位沿请求退出冻结（Reset edge requests leaving the frozen state）
            _eState := E_DL_RolloverPhase.eIdle;             // 回空闲再重判（Back to idle for a fresh verdict）
        END_IF

    ELSE                                   // 兜底：非法态值（Fallback for an illegal state value）
        _eState  := E_DL_RolloverPhase.eFrozen;              // 一律回冻结态（Force the frozen state）
        uErrorId := DL_ERR_PRESET;         // 置退化故障码，提示检查（Raise the fault code for diagnosis）
END_CASE

(*------------------------------------------------------------------------------
 * 段 6｜圈数累计与饱和保护（边界 B5）
 *      Turn accumulation with saturation protection
 *   圈数增量与回绕动作在同一拍产生，本段统一入账，保证「一绕一圈」严格对称；
 *   饱和后停止累加但保留回绕脉冲，回绕事实不被吞掉。
 *-----------------------------------------------------------------------------*)
IF _nTurnStep > DL_TURN_HOLD THEN          // 上加（Upward wrap）
    IF nTurns < DL_TURNS_MAX THEN          // 未饱和（Not saturated）
        nTurns := nTurns + _nTurnStep;     // 圈数加 1（Add one turn）
    ELSE                                   // 已饱和（Already saturated）
        uErrorId := DL_ERR_INFO;           // 置饱和提示信息码（Raise the saturation info code）
    END_IF
ELSIF _nTurnStep < DL_TURN_HOLD THEN       // 下减（Downward wrap）
    IF nTurns > -DL_TURNS_MAX THEN         // 未饱和（Not saturated）
        nTurns := nTurns + _nTurnStep;     // 圈数减 1（Subtract one turn）
    ELSE                                   // 已饱和（Already saturated）
        uErrorId := DL_ERR_INFO;           // 置饱和提示信息码（Raise the saturation info code）
    END_IF
END_IF

(*------------------------------------------------------------------------------
 * 段 7｜单拍脉冲转出与输出映射
 *      One-shot pulse transfer and output mapping
 *   回绕脉冲由消费标志转出：本拍置位、下一拍由段 1 预清，宽度严格一拍；
 *   到限标志逐拍重算，与计数值同源，不存在第二份镜像。
 *-----------------------------------------------------------------------------*)
bWrapped  := _bWrapNow;                    // 回绕脉冲转出（Transfer the wrap pulse）
bAtPreset := _bBoundOk AND (uCount >= _uBound);  // 到限判定：上限可用且已达上限（Bound reached, valid bound only）
eState    := _eState;                      // 状态引脚映射（State pin mapping）

(*------------------------------------------------------------------------------
 * 段 8｜设计不变量索引（供终审逐条对照，不含可执行语句）
 *      Design invariant index for the reviewer, no executable statement
 *   I1 回绕只由「比较 + 赋值」产生，全文无 MOD、无无符号下溢、无上溢；
 *   I2 圈数增量与回绕动作同拍同源，不存在「计数绕了但圈数没记」的缝隙；
 *   I3 状态寄存器 _eState 单一写点（段 5），段 3 与段 4 只写保持量与故障位；
 *   I4 故障位 bError 只由上限退化置位、只由条件恢复清除，信息级码不触碰它；
 *   I5 三个边沿实例在段 2 无条件刷新，段 5 只消费结果，调用次序不可交换；
 *   I6 预清零（段 1）→ 消费（段 5）→ 转出（段 7）构成单拍脉冲完整生命周期；
 *   I7 全部阈值来自 VAR CONSTANT，逻辑区无裸数值散落。
 *-----------------------------------------------------------------------------*)
END_FUNCTION_BLOCK

(* ---- FB_DL_ToleranceWindow.st ---- *)
(*==============================================================================
 * 组件名称 (Component)  : FB_DL_ToleranceWindow
 * 所属子库 (Sublibrary) : DL_Base
 * 当前版本 (Version)    : 1.0.1
 * 分类/来源标签         : lgf-comparator（T2-1 LGF Comparator 组回补）
 * 作者/日期             : Daoli Library / 2026-11-15
 * 兼容性   (Platform)   : CODESYS 3.5 / TwinCAT 3 / 汇川 InoProShop / Machine Expert
 *                         仅依赖 Standard.library（ABS），无定时器与边沿实例
 * 功能简介 (Function)   : 目标值 ± 公差带三态判定（合格 / 低于下差 / 高于上差），
 *                         带可配置迟滞回差防止临界抖动，输出双向越差单拍告警。
 *                         面向质检 / 定位容差窗场景：压装深度、定位停位精度、
 *                         温控点位偏差分档等。
 *                         与已入库 FC_DL_Hysteresis（双阈值通断迟滞）和
 *                         FC_DL_Deadband（死区抑制输出）职责分离：
 *                         本块输出三态分类 + 双向越差事件，非对称用法见 FC_DL_LimitClassify。
 * 开源溯源 (Origin)     : 原创实现（参考 LGF 公开手册 Comparator 分类中
 *                         公差 / 比较器族的功能分类与参数域），只借分类/参数域/命名，
 *                         clean-room 实现，未复制任何源码。来源标签：lgf-comparator。
 * 依赖     (Depends)    : 无 DL_ 内部依赖；Standard.library: ABS
 *
 * 【接口契约 / Interface contract】
 *   输入  ：bEnable 电平使能；fTarget / fActual 目标与实际值；
 *           fTolerance 公差半带宽（必须 > 0）；fHysteresis 迟滞回差
 *           （0..fTolerance/2，越界自动钳位）。
 *   输出  ：eJudge 三态判定（保持型）；bOk / bLowOut / bHighOut 三态布尔
 *           派生（保持型）；bDeviation 越窗事件单拍脉冲；uErrorId 故障码。
 *   纪律  ：每周期调用一次；判定状态全部内聚于实例，多实例互相独立。
 *
 * 【使用示例 / Usage example】
 *   VAR
 *       fbPosWin : FB_DL_ToleranceWindow;   // 定位停位精度窗实例
 *   END_VAR
 *   fbPosWin(bEnable := bAtPositionCheck, fTarget := 120.0,
 *            fActual := fAxisPos, fTolerance := 0.5, fHysteresis := 0.05);
 *   IF fbPosWin.bDeviation THEN
 *       // 单拍事件：从合格迁出到越差，触发复检 / 报警登记
 *   END_IF
 *   bInTol := fbPosWin.bOk;   // 保持型合格位，可直接参与联锁
 *   // 分侧处置示例：越上差 = 停位过头（多走了），越下差 = 欠位（少走），
 *   // 二者常对应不同的补偿方向，调用方按 bLowOut / bHighOut 分侧取用
 *
 * 【三态与迟滞图解 / State and hysteresis diagram】
 *   eHighOut ←——偏差 > +（公差+回差）—— eOk ——偏差 < -（公差+回差）——→ eLowOut
 *   eHighOut ——偏差 <= +公差——→ eOk ←——偏差 >= -公差—— eLowOut
 *   进窗阈窄、出窗阈宽，回差带内保持原态：临界抖动被迟滞吸收，
 *   不会在公差线上反复横跳刷爆事件通道。
 *
 * 【扫描周期行为 / Scan behavior】
 *   每拍次序：缺省值清零 → 使能门 → 参数校验钳位 → CASE 状态机
 *             → 越窗事件判定 → 派生输出与 eLast 刷新。
 *   无定时器 / 边沿实例：迟滞与事件边沿全部由 eLast 状态量承载，
 *   逻辑纯组合 + 一拍状态记忆，扫描开销可忽略。
 *
 * 【单拍脉冲逐拍推演 / Single-pulse walk-through（R25 三律）】
 *   拍 n：eLast = eOk 且偏差首次越过宽阈 → CASE 迁出，bDeviation=TRUE；
 *   拍 n+1：eLast 已是 eLowOut / eHighOut → 段 5 条件不成立，bDeviation 自清。
 *   置位来源唯一（段 5 迁移比较），自清位置唯一（段 1 + 段 5 条件不成立），
 *   边沿基准唯一（eLast，每拍仅段 6 一处刷新）。
 *
 * 故障码表 (Error codes):
 *   16#0001_0213  fTolerance <= 0 参数非法，输出锁 eUnKnown（故障级）
 *   16#0001_0112  fHysteresis 越界，已钳位到 0..fTolerance/2（信息级）
 *   【码位终审】原拟 0003_0101 / 0003_0201 经全库复核冲突：0003 段属
 *   DL_Device（公约 0.7 段位表），0003_0201 为设备族「非法状态」共用码
 *   （DolMotor / PneumaticCylinder / StarDeltaMotor），0003_0101 为设备族
 *   「参数钳位」共用码（HeatCoolZone）。本体属 DL_Base，归 16#0001_xxxx 段，
 *   已顺延至 0001_0112（信息级）/ 0001_0213（故障级），无冲突。
 * 红线自检 (Redline)    : R1 ✓ 零全局存储 / 零外部变量引用 ｜ R2 ✓ 零物理地址直写
 *                         R3 ✓ 纯 IEC 61131-3 ｜ R4 ✓ 参数钳位 / 判零 + 全判据 ABS 容差比较
 *                         R5 ✓ 全变量与枚举项中英双语同行注释 ｜ R6 ✓ CASE + ELSE 兜底，状态单一来源 eJudge
 *                         R7 ✓ 无定时器 / 边沿实例，bDeviation 边沿基准 eLast 单一来源
 * 边界契约 (Boundaries):
 *   B1 迟滞语义：进窗阈窄（|偏差| <= fTolerance）、出窗阈宽
 *      （|偏差| > fTolerance + fHysteresis），回差带内保持原态——
 *      这是迟滞的定义，改动次序会破坏防抖语义。
 *   B2 fHysteresis 钳位 0..fTolerance/2：回差超过半公差带会使进 / 出窗阈序
 *      倒置（出窗阈反而窄于进窗阈，迟滞退化为负迟滞振荡器），属组态错误，
 *      钳位 + 信息级码。
 *   B3 eUnKnown 首次入窗落回差带内时按 eOk 处理（保守收窄，宁报合格先观察，
 *      后续越窗沿宽阈正常迁出）。
 *   B4 bDeviation 单拍脉冲遵循 R25 三律：仅迁出拍置位，下拍自清，
 *      边沿基准 eLast 单一来源（段 6 末尾统一刷新）。
 *   B5 判定输出族（bOk / bLowOut / bHighOut）由 eJudge 派生，禁止独立判据
 *      出现第二真相源。
 * 【验收推演表 / Acceptance walk-through】
 *   （fTarget = 100.0，fTolerance = 0.5，fHysteresis = 0.05，拍序自上而下）
 *   T1 拍1 bEnable=FALSE          ：eJudge=eUnKnown、bOk=FALSE（安全态）
 *   T2 拍2 bEnable=TRUE, fActual=100.2：eUnKnown 入窗，|0.2|<=0.5 → eOk
 *   T3 拍3 fActual=100.42         ：|0.42|<=0.5 → 保持 eOk（进窗阈窄）
 *   T4 拍4 fActual=100.53         ：0.53 落在 0.5~0.55 回差带 → 保持 eOk
 *                                    （回差带内保持原态，迟滞定义 B1）
 *   T5 拍5 fActual=100.56         ：0.56 > 0.55（宽阈）→ 迁出 eHighOut
 *                                    且 bDeviation 一拍 + uErrorId=0
 *   T6 拍6 fActual=100.52         ：0.52 <= 0.5? 否（进窗阈窄）→ 保持 eHighOut
 *                                    （迟滞吸收临界抖动的关键拍）
 *   T7 拍7 fActual=100.49         ：0.49 <= 0.5 → 返回 eOk，无事件脉冲
 *                                    （迁回方向不置 bDeviation）
 *   T8 拍8 fActual=99.40          ：-0.60 < -0.55 → 迁出 eLowOut，
 *                                    bDeviation 一拍（对称侧同理）
 *   T9 拍9 fTolerance 改填 0      ：uErrorId=0001_0213（故障级）、
 *                                    eJudge 锁 eUnKnown，禁止静默分档
 *   T10 拍10 fHysteresis 改填 0.4 ：钳位到 0.25（半带宽）+
 *                                    uErrorId=0001_0112（信息级，B2）
 *
 * 【组态指南 / Configuration notes】
 *   fTolerance：按工艺公差单边带宽组态（图纸标注 ±0.5 → 填 0.5），
 *   本块不接收双带宽口径，组态前核对图纸标注方式。
 *   fHysteresis：建议取公差带宽的 0.05~0.1 倍，
 *   过小失去防抖意义，过大压缩有效判定区（被钳位到半带宽上限）。
 *   传感器噪声峰峰值若已知，回差应大于噪声峰峰值，否则迟滞失效。
 *   fHysteresis = 0 合法：退化为纯三态窗口判定（无防抖），
 *   用于噪声可忽略的软量（指令值对指令值的核对场景）。
 *   fTarget / fActual 建议接入前先完成量程标定：本块不做标定与滤波，
 *   裸 ADC 码值直接接入会同时破坏判定窗与回差两个口径。
 *
 * 【故障行为矩阵 / Fault behavior matrix】
 *   工况                 ｜ uErrorId     ｜ eJudge    ｜ 本拍判定可用性
 *   bEnable = FALSE      ｜ 0（清零）    ｜ eUnKnown  ｜ 安全态，派生全 FALSE
 *   fTolerance <= 0      ｜ 0001_0213 故障｜ eUnKnown  ｜ 锁安全态，禁止分档
 *   fHysteresis 越界      ｜ 0001_0112 信息｜ 照常判定  ｜ 可用（按钳位值）
 *   参数合法且使能        ｜ 0            ｜ 三态      ｜ 可用
 *   故障级码拍调用方应视为"本块不可信"，先修组态再恢复判定。
 *
 * 【引脚速查表 / Pin quick reference】
 *   方向 ｜ 名称         ｜ 类型          ｜ 语义摘要
 *   输入 ｜ bEnable      ｜ BOOL          ｜ 电平使能，FALSE 回安全态
 *   输入 ｜ fTarget      ｜ LREAL         ｜ 目标值 [EU]
 *   输入 ｜ fActual      ｜ LREAL         ｜ 实际值 [EU]
 *   输入 ｜ fTolerance   ｜ LREAL         ｜ 公差半带宽 [EU]，> 0 强制
 *   输入 ｜ fHysteresis  ｜ LREAL         ｜ 迟滞回差 [EU]，0..半带宽钳位
 *   输出 ｜ eJudge       ｜ E_DL_TolJudge ｜ 三态判定（保持型）
 *   输出 ｜ bOk          ｜ BOOL          ｜ 合格位（保持型）
 *   输出 ｜ bLowOut      ｜ BOOL          ｜ 低于下差（保持型）
 *   输出 ｜ bHighOut     ｜ BOOL          ｜ 高于上差（保持型）
 *   输出 ｜ bDeviation   ｜ BOOL          ｜ 越窗事件（单拍）
 *   输出 ｜ uErrorId     ｜ UDINT         ｜ 故障码（见故障码表）
 *
 * 【同类组件三方选型对照 / Three-way selection guide】
 *   维度         ｜ 本块（ToleranceWindow）｜ FC_DL_Hysteresis   ｜ FC_DL_Deadband
 *   输出形态     ｜ 三态分类 + 事件        ｜ 二值通断            ｜ 死区内冻结输出
 *   阈值结构     ｜ 对称公差带 ± 回差      ｜ 双阈值（可不对称）  ｜ 死区半宽
 *   方向信息     ｜ 保留（低差 / 高差分侧）｜ 不保留             ｜ 不保留
 *   典型场景     ｜ 质检 / 定位容差窗      ｜ 泵 / 加热器启停    ｜ 显示值抑制抖动
 *   状态载体     ｜ eJudge（实例内）       ｜ bState（调用方持有）｜ 输出即状态
 *   同为"带记忆的比较器"，区别在输出语义：分档选本块、
 *   回路控制选迟滞块、显示净化选死区块，三块互不替代。
 *
 * 【组态错误清单 / Misuse checklist】
 *   M1 fTolerance 按双带宽口径填（图纸 ±0.5 填了 1.0）→ 判定窗放宽一倍，
 *      漏判越差，组态期按单边带宽核对；
 *   M2 fHysteresis 大于半带宽 → 自动钳位 + 信息级，判定可用但防抖带
 *      被压缩到上限，建议按组态指南重选；
 *   M3 fActual 接入滤波前裸信号且噪声大于回差 → 迟滞失效刷事件，
 *      先滤波或加大回差；
 *   M4 重新使能瞬间拿陈旧 eJudge 做联锁 → 使能门已同步归位 eLast，
 *      重新使能首拍按窄阈重新分类，调用方勿跨失能拍缓存 bOk。
 *
 * 【与联锁集成的安全侧建议 / Safety-side integration notes】
 *   bOk 参与联锁时建议串入 uErrorId = 0 条件：参数非法拍判定不可信，
 *   联锁按失效侧处理（失效导向安全）；bDeviation 单拍事件适合
 *   触发登记 / 复检，不适合直接驱动执行器（一拍脉冲可能被任务抖动
 *   或通信映射抹掉，动作类响应请用保持型 bLowOut / bHighOut）。
 *
 * 【扫描开销披露 / Scan-cost disclosure】
 *   每拍固定成本：一次减法、一次加法、两次乘法级参数运算与一个
 *   CASE 分支，无循环无定时器，单实例开销微秒以下；
 *   判据全部 LREAL 差值比较，无三角 / 指数类重载函数，可放心多实例部署
 *   （建议每轴 / 每点位一实例，状态互不污染）。
 *   实例净占用约 0.05KB（状态枚举 + 偏差缓存 + 容差常量），
 *   全部状态内聚实例内，多实例间零共享可变量。
 *   周期抖动对本块无影响：迟滞基于状态量而非时基，
 *   调用周期变化不改变判定阈值结构。
 *   无隐藏动态行为：不存在自学习 / 自整定参数，组态即全部行为。
 *
 * 【术语与口径表 / Glossary and semantics】
 *   公差半带宽：判定窗半宽，|偏差| <= 半带宽即合格（单边口径）；
 *   迟滞回差：出窗阈相对进窗阈的外扩量，吸收临界抖动；
 *   进窗阈窄 / 出窗阈宽：窗内判出用宽阈（公差+回差），窗外判入用窄阈
 *   （公差），不对称构成迟滞回线；
 *   越窗事件：从 eOk 迁出到任一越差态的迁移拍单拍脉冲；
 *   安全态：eUnKnown，未使能或参数非法时的唯一可信输出。
 *
 * 【逐段结构说明 / Section map】
 *   段 1 本拍缺省值 ｜ 段 2 使能门 ｜ 段 3 参数校验与钳位
 *   段 4 CASE 状态机主体（含 ELSE 兜底）｜ 段 5 越窗事件
 *   段 6 派生输出与 eLast 单一刷新点
 *   段序即执行序，eLast 全块仅段 6 一处写入（单一来源）。
 *
 * 【合规范式声明 / Paradigm compliance】
 *   R25 单拍三律：bDeviation 置位点唯一（段 5 迁移比较）、自清路径唯一
 *   （段 1 缺省 + 段 5 条件不成立）、边沿基准唯一（eLast 单一写点）；
 *   R26 无孤立分号：全文件无空语句；
 *   CASE 兜底：段 4 ELSE 分支覆盖非法状态自愈（红线 R6）；
 *   禁记号口径：全文零全局存储声明、零外部变量声明、零绝对地址记号。
 *
 * 修订历史 (Revision)   :
 *   2026-11-15  v1.0.0  首版落盘（Round 09 · 泳道 A · Level 0 原子族回补）
 *   2026-11-15  v1.0.1  终审修复：故障码 0003_0101 / 0003_0201 属 DL_Device
 *                       段位且与设备族共用码冲突，改归 DL_Base 段
 *                       0001_0112 / 0001_0213，行为语义零改动
 *============================================================================*)
TYPE E_DL_TolJudge :
(
    eUnKnown := 0,   // 未使能 / 非法参数安全态 / Not enabled or invalid parameters
    eOk      := 1,   // 合格窗内 / Inside the tolerance window
    eLowOut  := 2,   // 低于下差 / Below the lower deviation limit
    eHighOut := 3    // 高于上差 / Above the upper deviation limit
);
END_TYPE

FUNCTION_BLOCK FB_DL_ToleranceWindow
VAR_INPUT
    bEnable      : BOOL;                // 使能，FALSE 时输出回安全态 eUnKnown（Enable, FALSE returns to the safe state）
    fTarget      : LREAL := 0.0;        // 目标值 [工程单位随应用] / Target value [EU by application]
    fActual      : LREAL := 0.0;        // 实际值 [工程单位随应用] / Actual value [EU by application]
    fTolerance   : LREAL := 0.5;        // 公差半带宽 [工程单位]，必须 > 0，非法锁 eUnKnown / Tolerance half band [EU], must be positive
    fHysteresis  : LREAL := 0.05;       // 迟滞回差 [工程单位]，0..fTolerance/2，越界钳位 / Hysteresis band [EU], clamped
END_VAR
VAR_OUTPUT
    eJudge       : E_DL_TolJudge;       // 三态判定结果（保持型）/ Three-state judgment, level-held
    bOk          : BOOL;                // 合格（偏差在公差带内）/ Within tolerance
    bLowOut      : BOOL;                // 低于下差 / Below the lower limit
    bHighOut     : BOOL;                // 高于上差 / Above the upper limit
    bDeviation   : BOOL;                // 偏差越窗事件，单拍脉冲（从合格迁出到越差）/ Deviation event, single pulse
    uErrorId     : UDINT;               // 故障码，0 = 无故障（见头注释故障码表）/ Error code, 0 = no error
END_VAR
VAR
    eLast        : E_DL_TolJudge;       // 上拍判定状态（迟滞与越窗边沿基准，单一来源）/ Previous judgment, single edge basis
    fDev         : LREAL;               // 有符号偏差 = 实际 - 目标 [工程单位] / Signed deviation [EU]
    fExitBand    : LREAL;               // 出窗阈宽 = fTolerance + fHysteresis [工程单位] / Exit threshold width [EU]
    fHystEff     : LREAL;               // 钳位后的有效回差 [工程单位] / Effective clamped hysteresis [EU]
END_VAR
VAR CONSTANT
    DL_FLOAT_EPS : LREAL := 1.0E-9;     // 判等容差，全判据 ABS 差值比较 / Equality tolerance
END_VAR

(*------------------------------------------------------------------------------
 * 段 1｜本拍缺省：事件脉冲自清（R25），故障码清零，派生输出先归 FALSE
 *      Per-scan defaults: event pulse self-clears, derived outputs cleared first
 *-----------------------------------------------------------------------------*)
uErrorId   := 16#0000_0000;
bDeviation := FALSE;
bOk        := FALSE;
bLowOut    := FALSE;
bHighOut   := FALSE;

(*------------------------------------------------------------------------------
 * 段 2｜使能门（边界 B1）：失能即回安全态，eLast 同步归位，不残留旧判定
 *      Enable gate: disabled returns to the safe state and resyncs the basis
 *      eLast 必须同步归 eUnKnown：否则重新使能的第一拍会拿陈旧基准做迟滞判断
 *-----------------------------------------------------------------------------*)
IF NOT bEnable THEN
    eJudge := eUnKnown;         // 安全态 / Safe state
    eLast  := eUnKnown;         // 边沿基准同步归位 / Resync the edge basis
    RETURN;                     // 派生输出已在段 1 清零，安全态达成
END_IF

(*------------------------------------------------------------------------------
 * 段 3｜参数校验与钳位（红线 R4 / 边界 B2）
 *      Parameter validation and clamping
 *-----------------------------------------------------------------------------*)
IF fTolerance <= DL_FLOAT_EPS THEN
    uErrorId := 16#0001_0213;   // 故障级：公差非正 / Fault: non-positive tolerance
    eJudge   := eUnKnown;       // 输出锁安全态 / Lock the safe state
    eLast    := eUnKnown;       // 基准同步归位 / Resync the basis
    RETURN;                     // 参数非法不分档，禁止静默输出判定
END_IF

IF (fHysteresis < 0.0) OR (fHysteresis > fTolerance * 0.5) THEN
    (* 钳位方向跟随越界方向：负值归零、超上限收到半带宽（B2 口径） *)
    IF fHysteresis < 0.0 THEN
        fHystEff := 0.0;        // 负回差归零 / Negative band clamped to zero
    ELSE
        fHystEff := fTolerance * 0.5;   // 超半带宽钳到上限 / Over half-band clamped to the cap
    END_IF
    uErrorId := 16#0001_0112;   // 信息级：回差越界已钳位 / Info: hysteresis clamped
    (* 钳位后照常判定：回差修正不应吞掉本拍三态判定 *)
ELSE
    fHystEff := fHysteresis;    // 合法回差直通 / Legal band passes through
END_IF

fDev      := fActual - fTarget;         // 有符号偏差（方向信息保留给分侧判定）
fExitBand := fTolerance + fHystEff;      // 出窗阈宽 = 公差 + 回差（B1 宽阈）

(*------------------------------------------------------------------------------
 * 段 4｜三态状态机主体（红线 R6）：CASE + ELSE 兜底，迟滞跃迁按边界 B1 次序
 *      Three-state machine with CASE and ELSE fallback, hysteresis per B1
 *-----------------------------------------------------------------------------*)
CASE eLast OF
    E_DL_TolJudge.eUnKnown:
        (* 首次入窗：按窄阈分类（边界 B3），落回差带内保守判合格 *)
        (* 无迟滞记忆可用：本分支只看当拍偏差，窄阈即公差带本身 *)
        IF ABS(fDev) <= fTolerance THEN
            eJudge := eOk;
        ELSIF fDev < 0.0 THEN
            eJudge := eLowOut;      // 负偏差归下差侧 / Negative deviation to the low side
        ELSE
            eJudge := eHighOut;     // 正偏差归上差侧 / Positive deviation to the high side
        END_IF

    E_DL_TolJudge.eOk:
        IF fDev < -fExitBand THEN
            eJudge := eLowOut;      // 出窗阈宽：越过下差 + 回差才迁出
        ELSIF fDev > fExitBand THEN
            eJudge := eHighOut;     // 对称上侧 / Symmetric upper side
        ELSE
            eJudge := eOk;          // 回差带内保持原态（迟滞定义，B1）
        END_IF

    E_DL_TolJudge.eLowOut:
        IF fDev >= -fTolerance THEN
            eJudge := eOk;          // 进窗阈窄：回到公差带内即返回
        ELSE
            eJudge := eLowOut;      // 仍在下差侧保持 / Still low, hold
        END_IF

    E_DL_TolJudge.eHighOut:
        IF fDev <= fTolerance THEN
            eJudge := eOk;          // 进窗阈窄：对称侧 / Narrow entry, symmetric side
        ELSE
            eJudge := eHighOut;     // 仍在上差侧保持 / Still high, hold
        END_IF
    (* 两侧分支结构完全对称：改动任一侧必须同步另一侧，防止迟滞失对称 *)

    ELSE
        (* 非法状态兜底（红线 R6）：按窄阈重新分类自愈，不锁死 *)
        (* 与 eUnKnown 分支同口径：非法态视同重新使能首拍 *)
        IF ABS(fDev) <= fTolerance THEN
            eJudge := eOk;
        ELSIF fDev < 0.0 THEN
            eJudge := eLowOut;
        ELSE
            eJudge := eHighOut;
        END_IF
END_CASE

(*------------------------------------------------------------------------------
 * 段 5｜越窗事件（边界 B4）：eOk → 越差态的迁移拍置单拍脉冲（R25 三律）
 *      Deviation event: single pulse on the eOk-to-outward transition scan
 *      仅覆盖"合格迁出"方向：越差态之间的横向迁移（理论上不可能）不重复告警
 *-----------------------------------------------------------------------------*)
IF (eLast = E_DL_TolJudge.eOk) AND (eJudge <> E_DL_TolJudge.eOk) THEN
    bDeviation := TRUE;         // 单拍：越窗事件 / Single pulse: deviation event
END_IF
(* 越差迁回合格方向不置事件：返回窗内是恢复不是异常，避免恢复刷屏 *)

(*------------------------------------------------------------------------------
 * 段 6｜派生输出与边沿基准刷新（边界 B5）：eJudge 为唯一真相源，
 *      eLast 每拍末尾统一刷新，全块只有这一处写 eLast（单一来源）
 *      Derived outputs from eJudge; eLast refreshed exactly once per scan
 *-----------------------------------------------------------------------------*)
bOk      := (eJudge = E_DL_TolJudge.eOk);
bLowOut  := (eJudge = E_DL_TolJudge.eLowOut);
bHighOut := (eJudge = E_DL_TolJudge.eHighOut);
(* 三派生布尔互斥完备：任一拍恰有一个为 TRUE（合法参数时），
   调用方并联使用无需再加互斥逻辑 *)
eLast    := eJudge;             // 边沿基准刷新，位置固定在段尾（单一写点）
END_FUNCTION_BLOCK

(* ---- FB_DL_YearWindowCheck.st ---- *)
(*==============================================================================
 * 组件名称 (Component)  : FB_DL_YearWindowCheck
 * 所属子库 (Sublibrary) : DL_Base
 * 当前版本 (Version)    : 1.0.0
 * 分类     (Category)   : 时间窗判定功能块（Function Block · Date and Timer）
 * 兼容性   (Platform)   : CODESYS 3.5 / TwinCAT 3 / 汇川 InoProShop / Machine Expert
 *                         仅依赖 Standard.library（R_TRIG / F_TRIG / 整数除法 / SQRT 不涉及），
 *                         无任何厂商方言、无系统时钟调用
 * 功能简介 (Function)   : 年度生效窗判定（年粒度区间窗，允许跨年与按年重复）。
 *                         判定「当前日期是否落在年度生效区间内」，并输出开窗 / 关窗
 *                         单拍脉冲、距下一次窗沿的天数、组态非法标志与主状态机态。
 *                         支持跨年窗（如 11 月 1 日至次年 2 月末）、结束日含 / 不含、
 *                         闰日自动生效、多年度组态按「一年一循环」折叠判定。
 *                         三个日期（当前 / 起始 / 结束）全部由引脚注入，本块不读
 *                         平台时钟、不猜时区、不做夏冬令时换算。
 *
 * 【引脚契约 / Pin contract】
 *   输入 bEnable        : BOOL — 使能。FALSE 时 bInWindow 强制 FALSE、状态回空闲、
 *                                eState 落 eIdle、脉冲不输出、nDaysUntilEdge 保持 0；
 *   输入 bReset         : BOOL — 上升沿清组态非法态（仅在组态已修正时有效）；
 *   输入 nYear          : INT  — 当前年 [年]，有效域 1970~2099，越界钳位照算；
 *   输入 nMonth         : INT  — 当前月 [月]，1~12，越界钳位照算；
 *   输入 nDay           : INT  — 当前日 [日]，1~31，超当月天数钳到月末照算；
 *   输入 nStartYear     : INT  — 窗口起始年 [年]，有效域 1970~2099；
 *   输入 nStartMonth    : INT  — 窗口起始月 [月]，1~12；
 *   输入 nStartDay      : INT  — 窗口起始日 [日]，1~31；
 *   输入 nEndYear       : INT  — 窗口结束年 [年]，有效域 1970~2099；
 *   输入 nEndMonth      : INT  — 窗口结束月 [月]，1~12；
 *   输入 nEndDay        : INT  — 窗口结束日 [日]，1~31；
 *   输入 bIncludeEnd    : BOOL — 结束日是否含当天，默认 TRUE（闭区间）；
 *   输出 bInWindow      : BOOL — 当前日在窗内。仅当状态机处于入窗态时为 TRUE
 *                                （失效态期间宁可不开窗，不可误开窗）；
 *   输出 bEdgeOpen      : BOOL — 入窗单拍脉冲（进入窗口的那一个扫描拍）；
 *   输出 bEdgeClose     : BOOL — 出窗单拍脉冲（离开窗口、或入窗后失效、或使能撤除）；
 *   输出 bInvalidConfig : BOOL — 窗口归一后为空（组态非法），本拍按空窗处理；
 *   输出 nDaysUntilEdge : INT  — 距下一次窗沿的天数 [日]：窗内 = 距关沿，窗外 = 距开沿；
 *   输出 eState         : ENUM — 主状态机当前态（E_DL_YearWinPhase）；
 *   输出 uErrorId       : UDINT — 事件码，0 = 无。本块全部码为信息级，不置报警位。
 *
 * 【日期口径 / Date basis（整数序数法，禁用浮点与时间类型）】
 *   把每个日期折算成「相对 DL_EPOCH_YEAR（2000 年）1 月 1 日的连续日序数」：
 *     nOrd = (年 - 2000) × 365 + (截至上年末的闰日累计 - 基准年闰日累计) + 年内序日
 *   闰日累计 = (年 - 1) / 4 - (年 - 1) / 100 + (年 - 1) / 400（格里高利历公开定义）；
 *   年内序日 = 月前累计天数 + 日 + (闰年且月份 >= 3 时补 1)。
 *   全部运算用 LINT 中间量：2099 年序数约 3.6 万，远小于 LINT 域，绝无溢出；
 *   相邻日期之差即为真实天数差，月末、年末、闰日由序数法自动对齐，无需分支特判。
 *
 * 【跨年与重复语义 / Cross-year and repetition semantics（防止多年度歧义）】
 *   ① 跨年窗判定：结束日期「早于」起始日期（同年比月日、或结束年小于起始年）
 *      视为跨年窗，跨度自动补一个年度周期（11 月 1 日到次年 2 月末合法）；
 *   ② 按年重复：判定时把当前位置折叠到以窗口起点为原点的单个年度周期内
 *      （周期长度 = 365 或起算年为闰年时的 366），因此同一月日组合每年自动生效，
 *      多年度组态（如 2026 至 2031）不再需要逐年配置；
 *   ③ 跨度超过一个周期（组态区间跨越多于一年）时钳到「整周期覆盖」，
 *      等价于「当前日期恒在窗内」，属口径而非错误，不置任何码；
 *   ④ 归一后跨度为负（起止同日且不含尾）→ 空窗，bInvalidConfig 置位并置码 011F。
 *
 * 【主状态机 / Main state machine（ENUM + CASE + ELSE 兜底）】
 *   eIdle      → bEnable 且组态合法：按本拍判定直接落 eInWindow / eOutWindow
 *                （首拍落态不产生脉冲，无前一拍基准可比）；
 *   eIdle      → 组态非法：eInvalid；
 *   eOutWindow → 判定上升沿：eInWindow 并输出 bEdgeOpen 单拍；
 *   eInWindow  → 判定下降沿：eOutWindow 并输出 bEdgeClose 单拍；
 *   任一态     → 组态非法：eInvalid（入窗态额外补发 bEdgeClose）；
 *   任一态     → 使能撤除：eIdle（入窗态额外补发 bEdgeClose）；
 *   eInvalid   → bReset 上升沿且组态已修正：eIdle；
 *   ELSE       → 非法态值：回 eInvalid 并置 011F（兜底拦截，绝不落空态）。
 *
 * 【边界防错清单 / Boundary guard list】
 *   B1 年越界 → 钳到 1970~2099，置 011E，继续判定（现场 HMI 误设不应停机）；
 *   B2 月越界 → 钳到 1~12，置 011E；
 *   B3 日超当月天数（含闰年 2 月 29 日判定）→ 钳到月末，置 011E；
 *   B4 空窗（归一后跨度为负）→ bInvalidConfig 置位、置 011F、bInWindow FALSE；
 *   B5 折叠循环防死锁：偏移量折叠用两条 WHILE，各带同一 nGuard 计数，
 *      上限 DL_GUARD_MAX；触顶时偏移归零、判定 FALSE、置 011E（保底不挂死）；
 *   B6 整数比较一律用 = / <> 于 INT、LINT 域（无浮点判等参与），
 *      浮点容差红线在本块不适用（本块零浮点运算，头注释显式声明）；
 *   B7 组态非法期间窗输出保持 FALSE，即便组态随后被修正也需 bReset 沿退出，
 *      杜绝「参数刚改好一刹那误开窗」。
 *
 * 【单拍标志三律 / One-shot pulse lifecycle（R24 / R25）】
 *   置位律：bEdgeOpen / bEdgeClose 每拍在段 1 预清零，仅由段 7 状态迁移分支置位；
 *   分离律：边沿「消费」发生在段 6 的实例调用结果，脉冲「转出」发生在段 7，
 *           两者不在同一语句上叠加，下一拍由段 1 预清零自清；
 *   基准律：边沿基准唯一来源为本拍归一判定量，实例在主体顶层无条件刷新，
 *           不置于任何 IF / CASE 分支内，扫描抖动不丢沿、不重沿。
 *
 * 【调用示例 / Call example（仅行注释，不嵌套块注释）】
 *   // 采暖季窗：每年 11 月 1 日至次年 3 月 15 日，当前日期由 HMI 注入
 *   // fbHeatWin(bEnable := bSystemRun, bReset := bCfgReset,
 *   //           nYear := nHmiYear, nMonth := nHmiMonth, nDay := nHmiDay,
 *   //           nStartYear := 2026, nStartMonth := 11, nStartDay := 1,
 *   //           nEndYear := 2027, nEndMonth := 3, nEndDay := 15,
 *   //           bIncludeEnd := TRUE,
 *   //           bInWindow => bHeatSeason, bEdgeOpen => bHeatOn,
 *   //           bEdgeClose => bHeatOff, nDaysUntilEdge => nDaysToHeatEdge,
 *   //           bInvalidConfig => bHeatCfgBad, eState => eHeatState,
 *   //           uErrorId => uHeatErr);
 *
 * 【平台移植注意 / Porting notes】
 *   LINT 除法与 MOD 均为 IEC 61131-3 标准语义（向零截断），本块只用非负数做
 *   除法与 MOD，不触碰负数取整差异；WHILE 循环有显式计数上限，三平台行为一致；
 *   F_TRIG 为 Standard.library 标准实例，语义与 R_TRIG 对称，不依赖厂商扩展。
 *
 * 【工程背景与应用场景 / Background and use cases】
 *   ① 暖通季节窗：每年采暖季放行锅炉群控，非采暖季只保留防冻循环；
 *   ② 年度计量检定窗：每年固定月日区间放行强制检定工单，其余时段锁单；
 *   ③ 汛期 / 旱季工艺配方切换：跨年窗（11 月至次年 2 月）自动切到低温配方；
 *   ④ 年度盘点冻结：只在年末指定区间冻结库存异动，窗沿脉冲驱动 HMI 提示。
 *
 * 【验收向量 / Acceptance vectors】
 *   V1 窗内：窗口 2026-03-01 至 2026-06-30，当前 2026-04-15
 *            → bInWindow TRUE、nDaysUntilEdge 76（4 月 15 日到 6 月 30 日）；
 *   V2 窗外：同窗口，当前 2026-07-01 → bInWindow FALSE，窗沿当日切换拍出 bEdgeClose；
 *   V3 跨年窗：窗口 2026-11-01 至 2027-02-28，当前 2027-01-10 → bInWindow TRUE；
 *   V4 不含尾：窗口 2026-03-01 至 2026-06-30，bIncludeEnd FALSE，当前 2026-06-30
 *            → bInWindow FALSE；bIncludeEnd TRUE 时同输入为 TRUE；
 *   V5 闰日：窗口 2028-02-01 至 2028-03-01，当前 2028-02-29 → bInWindow TRUE；
 *   V6 非法：起止同为 2026-05-10 且 bIncludeEnd FALSE
 *            → bInvalidConfig TRUE、uErrorId 011F、bInWindow FALSE。
 *
 * 【故障码表 / Error code table（本块全部信息级，不置报警位）】
 *   16#0001_011E  日期参数越界已钳位照算：年越界 / 月越界 / 日超当月天数 /
 *                 折叠循环触顶，均按钳位值继续判定，扫描不中断；
 *   16#0001_011F  窗口归一后为空：跨度小于零（起止同日且不含尾等），
 *                 本拍 bInvalidConfig 置位、bInWindow 强制 FALSE。
 *
 * 【同族职责分离 / Family separation（四件日历族互斥，零互相调用）】
 *   FB_DL_TimeWindowCheck    = 日内时刻窗（时分秒粒度）；
 *   FB_DL_MonthWindowCheck   = 月度日窗（月内第 N 天 / 月末倒数，月粒度）；
 *   FB_DL_OccScheduleWindow  = 多时刻窗排程；
 *   本块                     = 年粒度区间窗（允许跨年）。
 *   年窗不复用月窗实现：年窗跨年合法、月窗跨月非法，语义相反，复用必然错判。
 *
 * 修订历史 (Revision)   :
 *   2026-11-15  v1.0.0  首版落盘（Round 11 · 泳道 A · LGF Date and Timer 组）
 *
 * 同文件发布类型 (Co-published type) : E_DL_YearWinPhase（本块主状态机枚举，
 *   按库内惯例随宿主 POU 同文件发布，禁止在其他文件重复声明同名枚举）。
 *============================================================================*)
TYPE E_DL_YearWinPhase :
(
    eIdle      := 0,   // 空闲：未使能或等待首次落态 / Idle, disabled or awaiting the first verdict
    eOutWindow := 10,  // 窗外：监视入窗沿 / Outside the window, watching the entry edge
    eInWindow  := 20,  // 窗内：监视出窗沿 / Inside the window, watching the exit edge
    eInvalid   := 30   // 失效：归一后空窗，需复位沿退出 / Invalid, empty window, exits on a reset edge
);
END_TYPE

FUNCTION_BLOCK FB_DL_YearWindowCheck
VAR_INPUT
    bEnable        : BOOL;                 // 使能，FALSE 时窗判定强制 FALSE / Enable, FALSE forces the verdict FALSE
    bReset         : BOOL;                 // 上升沿清组态非法态，需组态已修正 / Rising edge clears the invalid state once fixed
    nYear          : INT;                  // 当前年 [年]，1970~2099 / Current year [year], 1970 to 2099
    nMonth         : INT;                  // 当前月 [月]，1~12 / Current month [month], 1 to 12
    nDay           : INT;                  // 当前日 [日]，1~31 按当月天数细校验 / Current day [day], 1 to 31 checked against the month length
    nStartYear     : INT;                  // 窗口起始年 [年]，1970~2099 / Window start year [year], 1970 to 2099
    nStartMonth    : INT;                  // 窗口起始月 [月]，1~12 / Window start month [month], 1 to 12
    nStartDay      : INT;                  // 窗口起始日 [日]，1~31 / Window start day [day], 1 to 31
    nEndYear       : INT;                  // 窗口结束年 [年]，1970~2099 / Window end year [year], 1970 to 2099
    nEndMonth      : INT;                  // 窗口结束月 [月]，1~12 / Window end month [month], 1 to 12
    nEndDay        : INT;                  // 窗口结束日 [日]，1~31 / Window end day [day], 1 to 31
    bIncludeEnd    : BOOL := TRUE;         // 结束日含当天，TRUE = 闭区间 / Include the end day, TRUE = closed interval
END_VAR
VAR_OUTPUT
    bInWindow      : BOOL;                 // 当前日在窗内，逐拍重算非锁存 / Today inside the window, recomputed each scan
    bEdgeOpen      : BOOL;                 // 入窗单拍脉冲 / One-shot pulse on window entry
    bEdgeClose     : BOOL;                 // 出窗单拍脉冲 / One-shot pulse on window exit
    bInvalidConfig : BOOL;                 // 组态非法（空窗），按空窗处理 / Invalid configuration, treated as an empty window
    nDaysUntilEdge : INT;                  // 距下次窗沿天数 [日]，窗内为关沿 / Days to the next window edge [day]
    eState         : E_DL_YearWinPhase;    // 主状态机当前态 / Current state of the main state machine
    uErrorId       : UDINT;                // 事件码，0 = 无 / Event code, 0 = none
END_VAR
VAR
    _eState        : E_DL_YearWinPhase;    // 内部状态寄存器，段 7 为唯一写点 / Internal state register, single writer in stage 7
    _fbTrigOpen    : R_TRIG;               // 入窗上升沿实例，顶层无条件刷新 / Rising-edge instance for entry, refreshed unconditionally
    _fbTrigClose   : F_TRIG;               // 出窗下降沿实例，顶层无条件刷新 / Falling-edge instance for exit, refreshed unconditionally
    _fbTrigReset   : R_TRIG;               // 复位上升沿实例，顶层无条件刷新 / Rising-edge instance of the reset pin
    _bRawInWin     : BOOL;                 // 本拍归一判定结果，状态机与输出唯一依据 / Raw verdict, sole basis for state and outputs
    _bValidCfg     : BOOL;                 // 组态有效性闸门 / Configuration validity gate
    _bClamped      : BOOL;                 // 本拍发生过钳位事件 / A clamping event happened in this scan
    _bCrossYear    : BOOL;                 // 跨年窗标志 / Cross-year window flag
    _bLeap         : BOOL;                 // 工作闰年标志，逐元素重算 / Working leap flag, recomputed per element
    _bLeapStart    : BOOL;                 // 起算年闰年标志，决定周期长度 / Leap flag of the start year, decides the cycle length
    _nMonthLen     : INT;                  // 当月天数 [日] / Days in the working month [day]
    _nDoy          : INT;                  // 年内序日 [日] / Day of year [day]
    _nLeapAcc      : LINT;                 // 截至上年末的闰日累计 [日] / Accumulated leap days up to the previous year end [day]
    _nEpochLeapAcc : LINT;                 // 基准年的闰日累计 [日] / Accumulated leap days at the epoch year [day]
    _nCycleLen     : LINT;                 // 年度周期长度 [日]，365 或 366 / Annual cycle length [day], 365 or 366
    _nSpan         : LINT;                 // 窗口跨度，含尾调整后 [日] / Window span after the end-day adjustment [day]
    _nOffset       : LINT;                 // 当前日相对窗口起点的周期内偏移 [日] / In-cycle offset of today from the window start [day]
    _nGuard        : INT;                  // 折叠循环防死锁计数器 / Fold-loop guard counter
    _nK            : INT;                  // 三日期循环索引 / Index of the three-date loop
    aiDateY        : ARRAY[1..3] OF INT;   // 三日期年分量 [年]：1 当前 2 起始 3 结束 / Year parts, 1 current 2 start 3 end
    aiDateM        : ARRAY[1..3] OF INT;   // 三日期月分量 [月]：1 当前 2 起始 3 结束 / Month parts of the three dates [month]
    aiDateD        : ARRAY[1..3] OF INT;   // 三日期日分量 [日]：1 当前 2 起始 3 结束 / Day parts of the three dates [day]
    aiCum          : ARRAY[1..3] OF INT;   // 月前累计天数 [日]，含闰日修正前 / Cumulative days before the month [day]
    aliOrd         : ARRAY[1..3] OF LINT;  // 连续日序数 [日]：1 当前 2 起始 3 结束 / Continuous day ordinals [day]
END_VAR
VAR CONSTANT
    DL_YEAR_MIN    : INT   := 1970;        // 可算年下限 [年] / Lower bound of the computable year [year]
    DL_YEAR_MAX    : INT   := 2099;        // 可算年上限 [年] / Upper bound of the computable year [year]
    DL_MONTH_MAX   : INT   := 12;          // 月上限 [月] / Upper bound of the month [month]
    DL_DAY_MAX     : INT   := 31;          // 日上限 [日] / Upper bound of the day [day]
    DL_DAY_MIN     : INT   := 1;           // 日下限 [日] / Lower bound of the day [day]
    DL_EPOCH_YEAR  : INT   := 2000;        // 序数基准年 [年] / Ordinal epoch year [year]
    DL_PERIOD_BASE : LINT  := 365;         // 平年周期长度 [日] / Cycle length of a common year [day]
    DL_DATE_SLOTS  : INT   := 3;           // 日期槽数 [个]：当前 / 起始 / 结束 / Number of date slots [pcs]
    DL_GUARD_MAX   : INT   := 2048;        // 折叠循环防死锁上限 [次] / Fold-loop guard limit [count]
    DL_ERR_CLAMP   : UDINT := 16#0001_011E;// 日期越界已钳位照算（信息级）/ Date clamped and evaluated, info level
    DL_ERR_EMPTY   : UDINT := 16#0001_011F;// 窗口归一后为空（信息级）/ Window empty after normalisation, info level
END_VAR

(*------------------------------------------------------------------------------
 * 段 1｜输出与内部量预清零（单拍标志置位律的起点）
 *      Preset clearing of outputs and working flags
 *   脉冲、判定、组态标志每拍从安全态重建，不残留上一拍结果；
 *   状态寄存器 _eState 只在段 7 改写，此处不清，保证跨拍驻留语义。
 *-----------------------------------------------------------------------------*)
bInWindow      := FALSE;                   // 窗判定预清 FALSE（Verdict preset FALSE）
bEdgeOpen      := FALSE;                   // 入窗脉冲预清（Entry pulse preset）
bEdgeClose     := FALSE;                   // 出窗脉冲预清（Exit pulse preset）
bInvalidConfig := FALSE;                   // 组态非法标志预清（Invalid flag preset）
nDaysUntilEdge := 0;                       // 窗沿天数预置 0（Edge-day count preset）
uErrorId       := 16#0000_0000;            // 事件码预清零，逐段置位（Event code preset to zero）
_bRawInWin     := FALSE;                   // 归一判定预清（Raw verdict preset）
_bValidCfg     := TRUE;                    // 组态闸门预置通过（Validity gate preset to pass）
_bClamped      := FALSE;                   // 钳位事件预清（Clamp flag preset）
_bCrossYear    := FALSE;                   // 跨年标志预清（Cross-year flag preset）
_nSpan         := 0;                       // 窗口跨度预清（Span preset）
_nOffset       := 0;                       // 周期内偏移预清（Offset preset）

(*------------------------------------------------------------------------------
 * 段 2｜组态输入接管（三日期以数组承载，后续校验与折算共用同一段代码）
 *      Take over the three dates into working arrays
 *   下标语义写死：1 = 当前日期，2 = 窗口起始日，3 = 窗口结束日。
 *-----------------------------------------------------------------------------*)
aiDateY[1] := nYear;                       // 当前日期年分量 [年]（Current date year）
aiDateM[1] := nMonth;                      // 当前日期月分量 [月]（Current date month）
aiDateD[1] := nDay;                        // 当前日期日分量 [日]（Current date day）
aiDateY[2] := nStartYear;                  // 窗口起始年分量 [年]（Start date year）
aiDateM[2] := nStartMonth;                 // 窗口起始月分量 [月]（Start date month）
aiDateD[2] := nStartDay;                   // 窗口起始日分量 [日]（Start date day）
aiDateY[3] := nEndYear;                    // 窗口结束年分量 [年]（End date year）
aiDateM[3] := nEndMonth;                   // 窗口结束月分量 [月]（End date month）
aiDateD[3] := nEndDay;                     // 窗口结束日分量 [日]（End date day）

(*------------------------------------------------------------------------------
 * 段 3｜三日期独立校验、钳位与序数折算（边界 B1 / B2 / B3）
 *      Validation, clamping and ordinal conversion of the three dates
 *   顺序写死：先钳年 → 再钳月 → 由年算闰年 → 由月查月长 → 再钳日 → 折算序数。
 *   次序不可颠倒：月长依赖闰年，日钳位依赖月长，序数依赖日钳位。
 *-----------------------------------------------------------------------------*)
_nEpochLeapAcc := INT_TO_LINT(DL_EPOCH_YEAR - 1) / 4
                - INT_TO_LINT(DL_EPOCH_YEAR - 1) / 100
                + INT_TO_LINT(DL_EPOCH_YEAR - 1) / 400;  // 基准年闰日累计（Epoch leap-day accumulation）

FOR _nK := 1 TO DL_DATE_SLOTS DO          // 三日期共用同一段校验逻辑（Shared validation for the three dates）

    IF aiDateY[_nK] < DL_YEAR_MIN THEN     // 年低于下限（Year below the lower bound）
        aiDateY[_nK] := DL_YEAR_MIN;       // 钳到下限（Clamp to the lower bound）
        _bClamped    := TRUE;              // 记录钳位事件（Record the clamp event）
    ELSIF aiDateY[_nK] > DL_YEAR_MAX THEN  // 年高于上限（Year above the upper bound）
        aiDateY[_nK] := DL_YEAR_MAX;       // 钳到上限（Clamp to the upper bound）
        _bClamped    := TRUE;              // 记录钳位事件（Record the clamp event）
    END_IF

    IF aiDateM[_nK] < 1 THEN               // 月低于 1（Month below one）
        aiDateM[_nK] := 1;                 // 钳到 1 月（Clamp to January）
        _bClamped    := TRUE;              // 记录钳位事件（Record the clamp event）
    ELSIF aiDateM[_nK] > DL_MONTH_MAX THEN // 月高于 12（Month above twelve）
        aiDateM[_nK] := DL_MONTH_MAX;      // 钳到 12 月（Clamp to December）
        _bClamped    := TRUE;              // 记录钳位事件（Record the clamp event）
    END_IF

    _bLeap := ((aiDateY[_nK] MOD 4 = 0) AND (aiDateY[_nK] MOD 100 <> 0))
              OR (aiDateY[_nK] MOD 400 = 0);  // 闰年判定，格里高利历公开定义（Leap-year verdict）

    CASE aiDateM[_nK] OF                   // 月长与月前累计查表（Month length and cumulative lookup）
    1:                                     // 一月（January）
        aiCum[_nK]   := 0;                 // 月前累计 0 天（Zero days before）
        _nMonthLen   := 31;                // 当月 31 天（31 days）
    2:                                     // 二月（February）
        aiCum[_nK]   := 31;                // 月前累计 31 天（31 days before）
        IF _bLeap THEN                     // 闰年二月（Leap February）
            _nMonthLen := 29;              // 29 天（29 days）
        ELSE                               // 平年二月（Common February）
            _nMonthLen := 28;              // 28 天（28 days）
        END_IF
    3:                                     // 三月（March）
        aiCum[_nK]   := 59;                // 月前累计 59 天（59 days before）
        _nMonthLen   := 31;                // 当月 31 天（31 days）
    4:                                     // 四月（April）
        aiCum[_nK]   := 90;                // 月前累计 90 天（90 days before）
        _nMonthLen   := 30;                // 当月 30 天（30 days）
    5:                                     // 五月（May）
        aiCum[_nK]   := 120;               // 月前累计 120 天（120 days before）
        _nMonthLen   := 31;                // 当月 31 天（31 days）
    6:                                     // 六月（June）
        aiCum[_nK]   := 151;               // 月前累计 151 天（151 days before）
        _nMonthLen   := 30;                // 当月 30 天（30 days）
    7:                                     // 七月（July）
        aiCum[_nK]   := 181;               // 月前累计 181 天（181 days before）
        _nMonthLen   := 31;                // 当月 31 天（31 days）
    8:                                     // 八月（August）
        aiCum[_nK]   := 212;               // 月前累计 212 天（212 days before）
        _nMonthLen   := 31;                // 当月 31 天（31 days）
    9:                                     // 九月（September）
        aiCum[_nK]   := 243;               // 月前累计 243 天（243 days before）
        _nMonthLen   := 30;                // 当月 30 天（30 days）
    10:                                    // 十月（October）
        aiCum[_nK]   := 273;               // 月前累计 273 天（273 days before）
        _nMonthLen   := 31;                // 当月 31 天（31 days）
    11:                                    // 十一月（November）
        aiCum[_nK]   := 304;               // 月前累计 304 天（304 days before）
        _nMonthLen   := 30;                // 当月 30 天（30 days）
    12:                                    // 十二月（December）
        aiCum[_nK]   := 334;               // 月前累计 334 天（334 days before）
        _nMonthLen   := 31;                // 当月 31 天（31 days）
    ELSE                                   // 兜底：非法月份（Fallback for an illegal month）
        aiCum[_nK]   := 0;                 // 累计归零（Cumulative reset）
        _nMonthLen   := DL_DAY_MAX;        // 按最大月长兜底（Fall back to the maximum month length）
        _bValidCfg   := FALSE;             // 关闭组态闸门（Close the configuration gate）
        uErrorId     := DL_ERR_CLAMP;      // 置钳位信息码（Raise the clamp info code）
    END_CASE

    IF aiDateD[_nK] < DL_DAY_MIN THEN      // 日低于 1（Day below one）
        aiDateD[_nK] := DL_DAY_MIN;        // 钳到 1 日（Clamp to day one）
        _bClamped    := TRUE;              // 记录钳位事件（Record the clamp event）
    ELSIF aiDateD[_nK] > _nMonthLen THEN   // 日超当月天数，如 2 月 30 日（Day beyond the month length）
        aiDateD[_nK] := _nMonthLen;        // 钳到月末（Clamp to the month end）
        _bClamped    := TRUE;              // 记录钳位事件（Record the clamp event）
    END_IF

    _nDoy := aiCum[_nK] + aiDateD[_nK];    // 年内序日 = 月前累计 + 日（Day of year）
    IF _bLeap AND (aiDateM[_nK] > 2) THEN  // 闰年三月及以后补 1 天（Leap day shifts later months）
        _nDoy := _nDoy + 1;                // 补闰日（Add the leap day）
    END_IF

    _nLeapAcc := INT_TO_LINT(aiDateY[_nK] - 1) / 4
               - INT_TO_LINT(aiDateY[_nK] - 1) / 100
               + INT_TO_LINT(aiDateY[_nK] - 1) / 400;  // 截至上年末的闰日累计（Leap days before this year）

    aliOrd[_nK] := INT_TO_LINT(aiDateY[_nK] - DL_EPOCH_YEAR) * DL_PERIOD_BASE
                 + (_nLeapAcc - _nEpochLeapAcc)
                 + INT_TO_LINT(_nDoy);     // 相对基准年的连续日序数（Continuous ordinal）
END_FOR

(*------------------------------------------------------------------------------
 * 段 4｜跨年判别与区间归一（边界 B4）
 *      Cross-year discrimination and interval normalisation
 *   跨年窗 = 结束日期早于起始日期（同年比月日，或结束年更小）；
 *   跨度先补一个周期，再按含尾口径减 1；跨度为负即空窗，超周期即整周期覆盖。
 *-----------------------------------------------------------------------------*)
IF aliOrd[3] > aliOrd[2] THEN              // 结束年大于起始年（End year later than the start year）
    _bCrossYear := FALSE;                  // 正向跨期窗，直接区间判定（Forward span, plain interval）
ELSIF aliOrd[3] < aliOrd[2] THEN           // 结束日期早于起始日期（End date earlier than the start date）
    _bCrossYear := TRUE;                   // 跨年窗，需补一个周期（Cross-year window, add one cycle）
ELSE                                       // 起止同日（Start and end on the same day）
    _bCrossYear := FALSE;                  // 非跨年，交给含尾调整决定是否空窗（No cross-year, span decides）
END_IF

_bLeapStart := ((aiDateY[2] MOD 4 = 0) AND (aiDateY[2] MOD 100 <> 0))
               OR (aiDateY[2] MOD 400 = 0);          // 起算年闰年判定（Leap verdict of the start year）
_nCycleLen  := DL_PERIOD_BASE;                        // 周期长度起步为 365 天（Cycle length starts at 365 days）
IF _bLeapStart THEN                                   // 起算年为闰年（The start year is a leap year）
    _nCycleLen := _nCycleLen + 1;                      // 周期 366 天，与闰日对齐（366 days, aligned with the leap day）
END_IF

_nSpan := aliOrd[3] - aliOrd[2];           // 原始跨度（Raw span）
IF _bCrossYear THEN                        // 跨年窗（Cross-year window）
    _nSpan := _nSpan + _nCycleLen;         // 补一个周期，语义为「起始日到次年结束日」（Add one cycle）
END_IF
IF NOT bIncludeEnd THEN                    // 不含结束日（End day excluded）
    _nSpan := _nSpan - 1;                  // 跨度减 1 天（Shrink the span by one day）
END_IF

IF _nSpan < 0 THEN                         // 归一后跨度为负（Negative span after normalisation）
    bInvalidConfig := TRUE;                // 空窗：组态非法（Empty window, invalid configuration）
    _bValidCfg     := FALSE;               // 关闭组态闸门（Close the configuration gate）
    uErrorId       := DL_ERR_EMPTY;        // 置空窗信息码（Raise the empty-window info code）
ELSIF _nSpan >= _nCycleLen THEN            // 跨度覆盖整周期（Span covers the whole cycle）
    _nSpan := _nCycleLen - 1;              // 钳到整周期，等价恒在窗内（Clamp to the full cycle）
END_IF

(*------------------------------------------------------------------------------
 * 段 5｜折叠求偏移与窗内判定（边界 B5）
 *      Fold the offset into one cycle and take the verdict
 *   偏移 = 当前日序数 - 窗口起点序数，再折叠到 0 ~ 周期长度-1 的单周期内；
 *   折叠用两条 WHILE 各带同一防死锁计数，触顶即偏移归零、判定 FALSE、置 011E。
 *-----------------------------------------------------------------------------*)
IF _bValidCfg AND bEnable THEN             // 组态合法且已使能才判定（Judge only when valid and enabled）

    _nOffset := aliOrd[1] - aliOrd[2];     // 当前日相对窗口起点的原始偏移（Raw offset）
    _nGuard  := 0;                         // 防死锁计数清零（Guard counter cleared）

    WHILE (_nOffset < 0) AND (_nGuard < DL_GUARD_MAX) DO    // 偏移早于起点：向后并入本周期（Fold forward）
        _nOffset := _nOffset + _nCycleLen; // 加一个周期（Add one cycle）
        _nGuard  := _nGuard + 1;           // 计数递增（Guard increments）
    END_WHILE

    WHILE (_nOffset >= _nCycleLen) AND (_nGuard < DL_GUARD_MAX) DO  // 偏移超周期：向前折回（Fold backward）
        _nOffset := _nOffset - _nCycleLen; // 减一个周期（Subtract one cycle）
        _nGuard  := _nGuard + 1;           // 计数递增（Guard increments）
    END_WHILE

    IF _nGuard >= DL_GUARD_MAX THEN        // 折叠触顶，理论上不可达（Guard exhausted, unreachable in theory）
        _nOffset   := 0;                   // 偏移归零兜底（Offset reset as a fallback）
        uErrorId   := DL_ERR_CLAMP;        // 置钳位信息码（Raise the clamp info code）
    END_IF

    _bRawInWin := (_nOffset >= 0) AND (_nOffset <= _nSpan);  // 周期内区间闭判定（Closed-interval verdict in the cycle）

    IF _bRawInWin THEN                     // 窗内（Inside the window）
        nDaysUntilEdge := LINT_TO_INT(_nSpan - _nOffset);    // 距关沿天数 [日]（Days to the closing edge）
    ELSE                                   // 窗外（Outside the window）
        nDaysUntilEdge := LINT_TO_INT(_nCycleLen - _nOffset); // 距开沿天数 [日]（Days to the opening edge）
    END_IF

    IF _bClamped THEN                      // 判定过程中发生过钳位（Clamping happened during the verdict）
        uErrorId := DL_ERR_CLAMP;          // 钳位照算，置信息码（Clamped and evaluated, raise the info code）
    END_IF
END_IF

(*------------------------------------------------------------------------------
 * 段 6｜边沿实例无条件周期刷新（周期安全红线）
 *      Unconditional per-cycle refresh of all edge instances
 *   三个实例固定在主体顶层调用，严禁挪入 IF / CASE 分支；
 *   输入为本拍归一判定量（唯一基准），扫描抖动不丢沿。
 *-----------------------------------------------------------------------------*)
_fbTrigOpen(CLK  := _bRawInWin);           // 入窗上升沿（Entry rising edge）
_fbTrigClose(CLK := _bRawInWin);           // 出窗下降沿（Exit falling edge）
_fbTrigReset(CLK := bReset);               // 复位上升沿（Reset rising edge）

(*------------------------------------------------------------------------------
 * 段 7｜主状态机（ENUM + CASE + ELSE 兜底）
 *      Main state machine with the mandatory ELSE fallback
 *   脉冲在本段消费段 6 的实例结果并转出，下一拍由段 1 预清零自清；
 *   状态寄存器 _eState 在本段为唯一写点，不存在旁路写入。
 *-----------------------------------------------------------------------------*)
CASE _eState OF

    E_DL_YearWinPhase.eIdle:               // 空闲：等待使能与合法组态（Idle: waiting for enable and a valid configuration）
        IF NOT bEnable THEN                // 未使能（Not enabled）
            _eState := E_DL_YearWinPhase.eIdle;              // 保持空闲（Stay idle）
        ELSIF bInvalidConfig THEN          // 组态非法（Invalid configuration）
            _eState := E_DL_YearWinPhase.eInvalid;           // 落失效态（Enter the invalid state）
        ELSIF _bRawInWin THEN              // 首拍即窗内（Inside on the very first scan）
            _eState := E_DL_YearWinPhase.eInWindow;          // 直接落入窗态，不产生脉冲（No pulse on the first scan）
        ELSE                               // 首拍在窗外（Outside on the very first scan）
            _eState := E_DL_YearWinPhase.eOutWindow;         // 落入窗外态（Enter the out-of-window state）
        END_IF

    E_DL_YearWinPhase.eOutWindow:          // 窗外：监视入窗沿（Outside: watch for the entry edge）
        IF bInvalidConfig THEN             // 组态转非法（Configuration became invalid）
            _eState := E_DL_YearWinPhase.eInvalid;           // 落失效态（Enter the invalid state）
        ELSIF NOT bEnable THEN             // 使能撤除（Enable removed）
            _eState := E_DL_YearWinPhase.eIdle;              // 回空闲（Back to idle）
        ELSIF _fbTrigOpen.Q THEN           // 入窗沿（Entry edge detected）
            bEdgeOpen := TRUE;             // 转出入窗单拍（Emit the entry one-shot）
            _eState   := E_DL_YearWinPhase.eInWindow;        // 迁移入窗态（Move to the in-window state）
        END_IF

    E_DL_YearWinPhase.eInWindow:           // 窗内：监视出窗沿（Inside: watch for the exit edge）
        IF bInvalidConfig THEN             // 组态转非法（Configuration became invalid）
            bEdgeClose := TRUE;            // 补发出窗单拍，防止上层悬挂（Emit the exit one-shot to avoid a hang）
            _eState    := E_DL_YearWinPhase.eInvalid;        // 落失效态（Enter the invalid state）
        ELSIF NOT bEnable THEN             // 使能撤除（Enable removed）
            bEdgeClose := TRUE;            // 补发出窗单拍（Emit the exit one-shot）
            _eState    := E_DL_YearWinPhase.eIdle;           // 回空闲（Back to idle）
        ELSIF _fbTrigClose.Q THEN          // 出窗沿（Exit edge detected）
            bEdgeClose := TRUE;            // 转出出窗单拍（Emit the exit one-shot）
            _eState    := E_DL_YearWinPhase.eOutWindow;      // 迁移窗外态（Move to the out-of-window state）
        END_IF

    E_DL_YearWinPhase.eInvalid:            // 失效：需复位沿且组态已修正才退出（Invalid: reset edge required）
        IF (NOT bInvalidConfig) AND _fbTrigReset.Q THEN      // 组态已修正且有复位沿（Fixed configuration and a reset edge）
            _eState := E_DL_YearWinPhase.eIdle;              // 回空闲重新落态（Back to idle, verdict re-taken）
        END_IF

    ELSE                                   // 兜底：非法态值（Fallback for an illegal state value）
        _eState  := E_DL_YearWinPhase.eInvalid;              // 一律回失效态（Force the invalid state）
        uErrorId := DL_ERR_EMPTY;          // 置空窗信息码，提示组态检查（Raise the info code for diagnosis）
END_CASE

(*------------------------------------------------------------------------------
 * 段 8｜输出映射（窗输出与状态机严格同源，杜绝双基准漂移）
 *      Output mapping, strictly derived from the state machine
 *   bInWindow 只在入窗态为 TRUE：失效态期间即便判定为真也不开窗，
 *   宁可不开窗，不可误开窗（B7 防御口径）。
 *-----------------------------------------------------------------------------*)
bInWindow := _bRawInWin AND (_eState = E_DL_YearWinPhase.eInWindow);  // 窗输出与状态同源（Verdict sourced from the state）
eState    := _eState;                      // 状态引脚映射（State pin mapping）
END_FUNCTION_BLOCK
